   "FRK_ConfigAppend"(Scope := #Scope,
                      Item := 'CatalogCount',
                      ValueText := WSTRING#'0',
                      ValueType := 0,
                      ReadLevel := #ReadLevel,
                      Readable := #Readable,
                      Cursor := #Cursor,
                      Page := #Page);
   "FRK_ConfigAppend"(Scope := #Scope,
                      Item := 'AvailableModelCount',
                      ValueText := INT_TO_WSTRING(#ModelCount),
                      ValueType := 0,
                      ReadLevel := #ReadLevel,
                      Readable := #Readable,
                      Cursor := #Cursor,
                      Page := #Page);
   FOR #Index := 0 TO 6 DO
       #IndexText := INT_TO_STRING(#Index);
       IF #IndexText[1] = '+' THEN
           #IndexText := DELETE(IN := #IndexText, L := 1, P := 1);
       END_IF;
       #Prefix := CONCAT(IN1 := 'ModePolicy/ModePolicy[', IN2 := #IndexText);
       #Prefix := CONCAT(IN1 := #Prefix, IN2 := ']/');
       #Item := CONCAT(IN1 := #Prefix, IN2 := 'Shield');
       "FRK_ConfigAppend"(Scope := #Scope,
                          Item := #Item,
                          ValueText := STRING_TO_WSTRING(DINT_TO_STRING(#Policy[#Index].Shield)),
                          ValueType := 0,
                          ReadLevel := #ReadLevel,
                          Readable := #Readable,
                          Cursor := #Cursor,
                          Page := #Page);
       #Item := CONCAT(IN1 := #Prefix, IN2 := 'Style');
       "FRK_ConfigAppend"(Scope := #Scope,
                          Item := #Item,
                          ValueText := STRING_TO_WSTRING(DINT_TO_STRING(#Policy[#Index].Style)),
                          ValueType := 0,
                          ReadLevel := #ReadLevel,
                          Readable := #Readable,
                          Cursor := #Cursor,
                          Page := #Page);
   END_FOR;
END_FUNCTION

FUNCTION "FRK_Config_DeclarationCell" : Void   // FC141, SCL
{ S7_Optimized_Access := 'TRUE' }
VERSION : 0.1
// stored: AutoNumber true, IsIECCheckEnabled false, SetENOAutomatically false, UDAEnableTagReadback false
   VAR_INPUT
      Access : "FRK_Access";
      RootIndex : Int;
      ModelIndex : UDInt;
   END_VAR
   VAR_IN_OUT
      Module : "FB_DeclarationCell";
      Cursor : "FRK_ConfigCursor";
      Page : "ST_ConfigPage";
   END_VAR
   VAR_TEMP
      Ok : Bool;
   END_VAR
BEGIN

   IF #ModelIndex = 0 THEN
       "FRK_ConfigCatalog"(Scope := #Module.Status.Name,
                           Catalog := #Module.Catalog,
                           Count := #Module.CatalogCount,
                           ReadLevel := #Access.Policy.Required[0],
                           Readable := #Access.CurrentLevel >= #Access.Policy.Required[0],
                           Cursor := #Cursor,
                           Page := #Page);
   END_IF;
   IF #ModelIndex = 0 THEN
       "FRK_CfgDef_DeclarationCell"(FieldIndex := 1);
       "FRK_ConfigScratch".Entry.Scope := STRING_TO_WSTRING(#Module.Status.Name);
       "FRK_ConfigScratch".Entry.ReadLevel := MAX(IN1 := #Access.Policy.Required[0], IN2 := "FRK_ConfigScratch".MinRead);
       "FRK_ConfigScratch".Entry.WriteLevel := MAX(IN1 := #Access.Policy.Required[1], IN2 := "FRK_ConfigScratch".MinWrite);
       "FRK_ConfigScratch".Entry.Readable := #Access.CurrentLevel >= "FRK_ConfigScratch".Entry.ReadLevel;
       "FRK_ConfigScratch".Entry.ModelScoped := FALSE;
       "FRK_ConfigScratch".Entry.ValueText := DINT_TO_WSTRING(TIME_TO_DINT(#Module.ParCfg.Timeout));
       IF NOT "FRK_ConfigScratch".Entry.Readable THEN
           "FRK_ConfigScratch".Entry.ValueText := WSTRING#'';
       END_IF;
       "FRK_ConfigAppendEntry"(Cursor := #Cursor,
                               Page := #Page);
   END_IF;
   IF #ModelIndex = 0 THEN
       "FRK_CfgDef_DeclarationCell"(FieldIndex := 2);
       "FRK_ConfigScratch".Entry.Scope := STRING_TO_WSTRING(#Module.Status.Name);
       "FRK_ConfigScratch".Entry.ReadLevel := MAX(IN1 := #Access.Policy.Required[0], IN2 := "FRK_ConfigScratch".MinRead);
       "FRK_ConfigScratch".Entry.WriteLevel := MAX(IN1 := #Access.Policy.Required[1], IN2 := "FRK_ConfigScratch".MinWrite);
       "FRK_ConfigScratch".Entry.Readable := #Access.CurrentLevel >= "FRK_ConfigScratch".Entry.ReadLevel;
       "FRK_ConfigScratch".Entry.ModelScoped := FALSE;
       "FRK_ConfigScratch".Entry.ValueText := DINT_TO_WSTRING(#Module.ParCfg.Preset);
       IF NOT "FRK_ConfigScratch".Entry.Readable THEN
           "FRK_ConfigScratch".Entry.ValueText := WSTRING#'';
       END_IF;
       "FRK_ConfigAppendEntry"(Cursor := #Cursor,
                               Page := #Page);
   END_IF;
   IF #ModelIndex = 0 THEN
       "FRK_Config_DeclarationCylinder"(Module := #Module.Clamp,
                                        Access := #Access,
                                        RootIndex := #RootIndex,
                                        ModelIndex := #ModelIndex,
                                        Cursor := #Cursor,
                                        Page := #Page);
   END_IF;
   IF #ModelIndex = 0 THEN
       "FRK_Config_DeclarationCylinder"(Module := #Module.Gate,
                                        Access := #Access,
                                        RootIndex := #RootIndex,
                                        ModelIndex := #ModelIndex,
                                        Cursor := #Cursor,
                                        Page := #Page);
   END_IF;
END_FUNCTION

FUNCTION "FRK_Config_DeclarationCylinder" : Void   // FC133, SCL
{ S7_Optimized_Access := 'TRUE' }
VERSION : 0.1
// stored: AutoNumber true, IsIECCheckEnabled false, SetENOAutomatically false, UDAEnableTagReadback false
   VAR_INPUT
      Access : "FRK_Access";
      RootIndex : Int;
      ModelIndex : UDInt;
   END_VAR
   VAR_IN_OUT
      Module : "FB_DeclarationCylinder";
      Cursor : "FRK_ConfigCursor";
      Page : "ST_ConfigPage";
   END_VAR
   VAR_TEMP
      Ok : Bool;
   END_VAR
BEGIN

   IF #ModelIndex = 0 THEN
       "FRK_ConfigCatalog"(Scope := #Module.Status.Name,
                           Catalog := #Module.Catalog,
                           Count := #Module.CatalogCount,
                           ReadLevel := #Access.Policy.Required[0],
                           Readable := #Access.CurrentLevel >= #Access.Policy.Required[0],
                           Cursor := #Cursor,
                           Page := #Page);
   END_IF;
   IF #ModelIndex = 0 THEN
       "FRK_CfgDef_DeclarationCylinder"(FieldIndex := 1);
       "FRK_ConfigScratch".Entry.Scope := STRING_TO_WSTRING(#Module.Status.Name);
       "FRK_ConfigScratch".Entry.ReadLevel := MAX(IN1 := #Access.Policy.Required[0], IN2 := "FRK_ConfigScratch".MinRead);
       "FRK_ConfigScratch".Entry.WriteLevel := MAX(IN1 := #Access.Policy.Required[1], IN2 := "FRK_ConfigScratch".MinWrite);
       "FRK_ConfigScratch".Entry.Readable := #Access.CurrentLevel >= "FRK_ConfigScratch".Entry.ReadLevel;
       "FRK_ConfigScratch".Entry.ModelScoped := FALSE;
       "FRK_ConfigScratch".Entry.ValueText := DINT_TO_WSTRING(TIME_TO_DINT(#Module.ParCfg.Timeout));
       IF NOT "FRK_ConfigScratch".Entry.Readable THEN
           "FRK_ConfigScratch".Entry.ValueText := WSTRING#'';
       END_IF;
       "FRK_ConfigAppendEntry"(Cursor := #Cursor,
                               Page := #Page);
   END_IF;
   IF #ModelIndex = 0 THEN
       "FRK_CfgDef_DeclarationCylinder"(FieldIndex := 2);
       "FRK_ConfigScratch".Entry.Scope := STRING_TO_WSTRING(#Module.Status.Name);
       "FRK_ConfigScratch".Entry.ReadLevel := MAX(IN1 := #Access.Policy.Required[0], IN2 := "FRK_ConfigScratch".MinRead);
       "FRK_ConfigScratch".Entry.WriteLevel := MAX(IN1 := #Access.Policy.Required[1], IN2 := "FRK_ConfigScratch".MinWrite);
       "FRK_ConfigScratch".Entry.Readable := #Access.CurrentLevel >= "FRK_ConfigScratch".Entry.ReadLevel;
       "FRK_ConfigScratch".Entry.ModelScoped := FALSE;
       "FRK_ConfigScratch".Entry.ValueText := DINT_TO_WSTRING(#Module.ParCfg.Preset);
       IF NOT "FRK_ConfigScratch".Entry.Readable THEN
           "FRK_ConfigScratch".Entry.ValueText := WSTRING#'';
       END_IF;
       "FRK_ConfigAppendEntry"(Cursor := #Cursor,
                               Page := #Page);
   END_IF;
END_FUNCTION

FUNCTION "FRK_Config_DeclarationUnit" : Void   // FC166, SCL
{ S7_Optimized_Access := 'TRUE' }
VERSION : 0.1
// stored: AutoNumber true, IsIECCheckEnabled false, SetENOAutomatically false, UDAEnableTagReadback false
   VAR_INPUT
      Access : "FRK_Access";
      RootIndex : Int;
      ModelIndex : UDInt;
   END_VAR
   VAR_IN_OUT
      Core : "FRK_Core";
      Status : "ST_ModuleStatus";
      ParCfg : "ST_DeclarationParCfg";
      ModePolicy : Array[0..6] of "ST_ModePolicy";
      AvailableModelCount : Int;
      StationCfg : "ST_UnitProbeStationCfg";
      Cell : "FB_DeclarationCell";
      Satellite : "FB_SatelliteUnit";
      Cursor : "FRK_ConfigCursor";
      Page : "ST_ConfigPage";
   END_VAR
   VAR_TEMP
      Ok : Bool;
   END_VAR
BEGIN

   IF #ModelIndex = 0 THEN
       "FRK_ConfigUnit"(Scope := #Status.Name,
                        Policy := #ModePolicy,
                        ModelCount := #AvailableModelCount,
                        ReadLevel := #Access.Policy.Required[0],
                        Readable := #Access.CurrentLevel >= #Access.Policy.Required[0],
                        Cursor := #Cursor,
                        Page := #Page);
   END_IF;
   IF #ModelIndex = 0 THEN
       "FRK_ConfigAppend"(Scope := #Status.Name,
                          Item := 'AvailableModels/AvailableModels[1]/ModelCode',
                          ValueText := WSTRING#'MODEL_A',
                          ValueType := 1,
                          ReadLevel := #Access.Policy.Required[0],
                          Readable := #Access.CurrentLevel >= #Access.Policy.Required[0],
                          Cursor := #Cursor,
                          Page := #Page);
       "FRK_ConfigAppend"(Scope := #Status.Name,
                          Item := 'AvailableModels/AvailableModels[2]/ModelCode',
                          ValueText := WSTRING#'MODEL_B',
                          ValueType := 1,
                          ReadLevel := #Access.Policy.Required[0],
                          Readable := #Access.CurrentLevel >= #Access.Policy.Required[0],
                          Cursor := #Cursor,
                          Page := #Page);
   END_IF;
   IF (#ModelIndex = 0 OR #Core.ParentIndex = 0) THEN
       "FRK_CfgDef_DeclarationUnit"(FieldIndex := 1);
       "FRK_ConfigScratch".Entry.Scope := STRING_TO_WSTRING(#Status.Name);
       "FRK_ConfigScratch".Entry.ReadLevel := MAX(IN1 := #Access.Policy.Required[0], IN2 := "FRK_ConfigScratch".MinRead);
       "FRK_ConfigScratch".Entry.WriteLevel := MAX(IN1 := #Access.Policy.Required[1], IN2 := "FRK_ConfigScratch".MinWrite);
       "FRK_ConfigScratch".Entry.Readable := #Access.CurrentLevel >= "FRK_ConfigScratch".Entry.ReadLevel;
       "FRK_ConfigScratch".Entry.ModelScoped := #Core.ParentIndex = 0;
       IF #ModelIndex <> 0 THEN
           "FRK_ConfigScratch".Entry.RequiresReady := "FRK_ConfigScratch".Entry.RequiresReady AND "FRK_ConfigModelCode"(RootIndex := #RootIndex, ModelIndex := #ModelIndex) = "FRK_ConfigStore".ActiveModels[#RootIndex];
           #Ok := "FRK_ConfigGet"(Scope := #Status.Name, ModelCode := "FRK_ConfigModelCode"(RootIndex := #RootIndex, ModelIndex := #ModelIndex));
           IF NOT #Ok THEN
               "FRK_ConfigScratch".Entry.Readable := FALSE;
           END_IF;
       ELSE
           "FRK_ConfigScratch".Entry.ValueText := DINT_TO_WSTRING(TIME_TO_DINT(#ParCfg.Timeout));
       END_IF;
       IF NOT "FRK_ConfigScratch".Entry.Readable THEN
           "FRK_ConfigScratch".Entry.ValueText := WSTRING#'';
       END_IF;
       "FRK_ConfigAppendEntry"(Cursor := #Cursor,
                               Page := #Page);
   END_IF;
   IF (#ModelIndex = 0 OR #Core.ParentIndex = 0) THEN
       "FRK_CfgDef_DeclarationUnit"(FieldIndex := 2);
       "FRK_ConfigScratch".Entry.Scope := STRING_TO_WSTRING(#Status.Name);
       "FRK_ConfigScratch".Entry.ReadLevel := MAX(IN1 := #Access.Policy.Required[0], IN2 := "FRK_ConfigScratch".MinRead);
       "FRK_ConfigScratch".Entry.WriteLevel := MAX(IN1 := #Access.Policy.Required[1], IN2 := "FRK_ConfigScratch".MinWrite);
       "FRK_ConfigScratch".Entry.Readable := #Access.CurrentLevel >= "FRK_ConfigScratch".Entry.ReadLevel;
       "FRK_ConfigScratch".Entry.ModelScoped := #Core.ParentIndex = 0;
       IF #ModelIndex <> 0 THEN
           "FRK_ConfigScratch".Entry.RequiresReady := "FRK_ConfigScratch".Entry.RequiresReady AND "FRK_ConfigModelCode"(RootIndex := #RootIndex, ModelIndex := #ModelIndex) = "FRK_ConfigStore".ActiveModels[#RootIndex];
           #Ok := "FRK_ConfigGet"(Scope := #Status.Name, ModelCode := "FRK_ConfigModelCode"(RootIndex := #RootIndex, ModelIndex := #ModelIndex));
           IF NOT #Ok THEN
               "FRK_ConfigScratch".Entry.Readable := FALSE;
           END_IF;
       ELSE
           "FRK_ConfigScratch".Entry.ValueText := DINT_TO_WSTRING(#ParCfg.Preset);
       END_IF;
       IF NOT "FRK_ConfigScratch".Entry.Readable THEN
           "FRK_ConfigScratch".Entry.ValueText := WSTRING#'';
       END_IF;
       "FRK_ConfigAppendEntry"(Cursor := #Cursor,
                               Page := #Page);
   END_IF;
   IF #ModelIndex = 0 THEN
       "FRK_CfgDef_DeclarationUnit"(FieldIndex := 3);
       "FRK_ConfigScratch".Entry.Scope := STRING_TO_WSTRING(#Status.Name);
       "FRK_ConfigScratch".Entry.ReadLevel := MAX(IN1 := #Access.Policy.Required[0], IN2 := "FRK_ConfigScratch".MinRead);
       "FRK_ConfigScratch".Entry.WriteLevel := MAX(IN1 := #Access.Policy.Required[1], IN2 := "FRK_ConfigScratch".MinWrite);
       "FRK_ConfigScratch".Entry.Readable := #Access.CurrentLevel >= "FRK_ConfigScratch".Entry.ReadLevel;
       "FRK_ConfigScratch".Entry.ModelScoped := FALSE;
       "FRK_ConfigScratch".Entry.ValueText := STRING_TO_WSTRING(#StationCfg.SiteLabel);
       IF NOT "FRK_ConfigScratch".Entry.Readable THEN
           "FRK_ConfigScratch".Entry.ValueText := WSTRING#'';
       END_IF;
       "FRK_ConfigAppendEntry"(Cursor := #Cursor,
                               Page := #Page);
   END_IF;
   IF #ModelIndex = 0 THEN
       "FRK_CfgDef_DeclarationUnit"(FieldIndex := 4);
       "FRK_ConfigScratch".Entry.Scope := STRING_TO_WSTRING(#Status.Name);
       "FRK_ConfigScratch".Entry.ReadLevel := MAX(IN1 := #Access.Policy.Required[0], IN2 := "FRK_ConfigScratch".MinRead);
       "FRK_ConfigScratch".Entry.WriteLevel := MAX(IN1 := #Access.Policy.Required[1], IN2 := "FRK_ConfigScratch".MinWrite);
       "FRK_ConfigScratch".Entry.Readable := #Access.CurrentLevel >= "FRK_ConfigScratch".Entry.ReadLevel;
       "FRK_ConfigScratch".Entry.ModelScoped := FALSE;
       "FRK_ConfigScratch".Entry.ValueText := STRING_TO_WSTRING(#StationCfg.LongText);
       IF NOT "FRK_ConfigScratch".Entry.Readable THEN
           "FRK_ConfigScratch".Entry.ValueText := WSTRING#'';
       END_IF;
       "FRK_ConfigAppendEntry"(Cursor := #Cursor,
                               Page := #Page);
   END_IF;
   IF #ModelIndex = 0 THEN
       "FRK_CfgDef_DeclarationUnit"(FieldIndex := 5);
       "FRK_ConfigScratch".Entry.Scope := STRING_TO_WSTRING(#Status.Name);
       "FRK_ConfigScratch".Entry.ReadLevel := MAX(IN1 := #Access.Policy.Required[0], IN2 := "FRK_ConfigScratch".MinRead);
       "FRK_ConfigScratch".Entry.WriteLevel := MAX(IN1 := #Access.Policy.Required[1], IN2 := "FRK_ConfigScratch".MinWrite);
       "FRK_ConfigScratch".Entry.Readable := #Access.CurrentLevel >= "FRK_ConfigScratch".Entry.ReadLevel;
       "FRK_ConfigScratch".Entry.ModelScoped := FALSE;
       IF #StationCfg.Enabled THEN
           "FRK_ConfigScratch".Entry.ValueText := WSTRING#'true';
       ELSE
           "FRK_ConfigScratch".Entry.ValueText := WSTRING#'false';
       END_IF;
       IF NOT "FRK_ConfigScratch".Entry.Readable THEN
           "FRK_ConfigScratch".Entry.ValueText := WSTRING#'';
       END_IF;
       "FRK_ConfigAppendEntry"(Cursor := #Cursor,
                               Page := #Page);
   END_IF;
   IF #ModelIndex = 0 THEN
       "FRK_Config_DeclarationCell"(Module := #Cell,
                                    Access := #Access,
                                    RootIndex := #RootIndex,
                                    ModelIndex := #ModelIndex,
                                    Cursor := #Cursor,
                                    Page := #Page);
   END_IF;
   IF #ModelIndex = 0 THEN
       "FRK_Config_SatelliteUnit"(Module := #Satellite,
                                  Access := #Access,
                                  RootIndex := #RootIndex,
                                  ModelIndex := #ModelIndex,
                                  Cursor := #Cursor,
                                  Page := #Page);
   END_IF;
END_FUNCTION

FUNCTION "FRK_Config_InnerUnit" : Void   // FC150, SCL
{ S7_Optimized_Access := 'TRUE' }
VERSION : 0.1
// stored: AutoNumber true, IsIECCheckEnabled false, SetENOAutomatically false, UDAEnableTagReadback false
   VAR_INPUT
      Access : "FRK_Access";
      RootIndex : Int;
      ModelIndex : UDInt;
   END_VAR
   VAR_IN_OUT
      Module : "FB_InnerUnit";
      Cursor : "FRK_ConfigCursor";
      Page : "ST_ConfigPage";
   END_VAR
   VAR_TEMP
      Ok : Bool;
   END_VAR
BEGIN

   IF #ModelIndex = 0 THEN
       "FRK_ConfigUnit"(Scope := #Module.Status.Name,
                        Policy := #Module.ModePolicy,
                        ModelCount := 0,
                        ReadLevel := #Access.Policy.Required[0],
                        Readable := #Access.CurrentLevel >= #Access.Policy.Required[0],
                        Cursor := #Cursor,
                        Page := #Page);
   END_IF;
   IF #ModelIndex = 0 THEN
       "FRK_CfgDef_InnerUnit"(FieldIndex := 1);
       "FRK_ConfigScratch".Entry.Scope := STRING_TO_WSTRING(#Module.Status.Name);
       "FRK_ConfigScratch".Entry.ReadLevel := MAX(IN1 := #Access.Policy.Required[0], IN2 := "FRK_ConfigScratch".MinRead);
       "FRK_ConfigScratch".Entry.WriteLevel := MAX(IN1 := #Access.Policy.Required[1], IN2 := "FRK_ConfigScratch".MinWrite);
       "FRK_ConfigScratch".Entry.Readable := #Access.CurrentLevel >= "FRK_ConfigScratch".Entry.ReadLevel;
       "FRK_ConfigScratch".Entry.ModelScoped := FALSE;
       "FRK_ConfigScratch".Entry.ValueText := DINT_TO_WSTRING(TIME_TO_DINT(#Module.ParCfg.Timeout));
       IF NOT "FRK_ConfigScratch".Entry.Readable THEN
           "FRK_ConfigScratch".Entry.ValueText := WSTRING#'';
       END_IF;
       "FRK_ConfigAppendEntry"(Cursor := #Cursor,
                               Page := #Page);
   END_IF;
   IF #ModelIndex = 0 THEN
       "FRK_CfgDef_InnerUnit"(FieldIndex := 2);
       "FRK_ConfigScratch".Entry.Scope := STRING_TO_WSTRING(#Module.Status.Name);
       "FRK_ConfigScratch".Entry.ReadLevel := MAX(IN1 := #Access.Policy.Required[0], IN2 := "FRK_ConfigScratch".MinRead);
       "FRK_ConfigScratch".Entry.WriteLevel := MAX(IN1 := #Access.Policy.Required[1], IN2 := "FRK_ConfigScratch".MinWrite);
       "FRK_ConfigScratch".Entry.Readable := #Access.CurrentLevel >= "FRK_ConfigScratch".Entry.ReadLevel;
       "FRK_ConfigScratch".Entry.ModelScoped := FALSE;
       "FRK_ConfigScratch".Entry.ValueText := DINT_TO_WSTRING(#Module.ParCfg.Preset);
       IF NOT "FRK_ConfigScratch".Entry.Readable THEN
           "FRK_ConfigScratch".Entry.ValueText := WSTRING#'';
       END_IF;
       "FRK_ConfigAppendEntry"(Cursor := #Cursor,
                               Page := #Page);
   END_IF;
   IF #ModelIndex = 0 THEN
       "FRK_CfgDef_InnerUnit"(FieldIndex := 3);
       "FRK_ConfigScratch".Entry.Scope := STRING_TO_WSTRING(#Module.Status.Name);
       "FRK_ConfigScratch".Entry.ReadLevel := MAX(IN1 := #Access.Policy.Required[0], IN2 := "FRK_ConfigScratch".MinRead);
       "FRK_ConfigScratch".Entry.WriteLevel := MAX(IN1 := #Access.Policy.Required[1], IN2 := "FRK_ConfigScratch".MinWrite);
       "FRK_ConfigScratch".Entry.Readable := #Access.CurrentLevel >= "FRK_ConfigScratch".Entry.ReadLevel;
       "FRK_ConfigScratch".Entry.ModelScoped := FALSE;
       "FRK_ConfigScratch".Entry.ValueText := STRING_TO_WSTRING(#Module.StationCfg.SiteLabel);
       IF NOT "FRK_ConfigScratch".Entry.Readable THEN
           "FRK_ConfigScratch".Entry.ValueText := WSTRING#'';
       END_IF;
       "FRK_ConfigAppendEntry"(Cursor := #Cursor,
                               Page := #Page);
   END_IF;
   IF #ModelIndex = 0 THEN
       "FRK_CfgDef_InnerUnit"(FieldIndex := 4);
       "FRK_ConfigScratch".Entry.Scope := STRING_TO_WSTRING(#Module.Status.Name);
       "FRK_ConfigScratch".Entry.ReadLevel := MAX(IN1 := #Access.Policy.Required[0], IN2 := "FRK_ConfigScratch".MinRead);
       "FRK_ConfigScratch".Entry.WriteLevel := MAX(IN1 := #Access.Policy.Required[1], IN2 := "FRK_ConfigScratch".MinWrite);
       "FRK_ConfigScratch".Entry.Readable := #Access.CurrentLevel >= "FRK_ConfigScratch".Entry.ReadLevel;
       "FRK_ConfigScratch".Entry.ModelScoped := FALSE;
       "FRK_ConfigScratch".Entry.ValueText := STRING_TO_WSTRING(#Module.StationCfg.LongText);
       IF NOT "FRK_ConfigScratch".Entry.Readable THEN
           "FRK_ConfigScratch".Entry.ValueText := WSTRING#'';
       END_IF;
       "FRK_ConfigAppendEntry"(Cursor := #Cursor,
                               Page := #Page);
   END_IF;
   IF #ModelIndex = 0 THEN
       "FRK_CfgDef_InnerUnit"(FieldIndex := 5);
       "FRK_ConfigScratch".Entry.Scope := STRING_TO_WSTRING(#Module.Status.Name);
       "FRK_ConfigScratch".Entry.ReadLevel := MAX(IN1 := #Access.Policy.Required[0], IN2 := "FRK_ConfigScratch".MinRead);
       "FRK_ConfigScratch".Entry.WriteLevel := MAX(IN1 := #Access.Policy.Required[1], IN2 := "FRK_ConfigScratch".MinWrite);
       "FRK_ConfigScratch".Entry.Readable := #Access.CurrentLevel >= "FRK_ConfigScratch".Entry.ReadLevel;
       "FRK_ConfigScratch".Entry.ModelScoped := FALSE;
       IF #Module.StationCfg.Enabled THEN
           "FRK_ConfigScratch".Entry.ValueText := WSTRING#'true';
       ELSE
           "FRK_ConfigScratch".Entry.ValueText := WSTRING#'false';
       END_IF;
       IF NOT "FRK_ConfigScratch".Entry.Readable THEN
           "FRK_ConfigScratch".Entry.ValueText := WSTRING#'';
       END_IF;
       "FRK_ConfigAppendEntry"(Cursor := #Cursor,
                               Page := #Page);
   END_IF;
   IF #ModelIndex = 0 THEN
       "FRK_Config_DeclarationCell"(Module := #Module.Cell,
                                    Access := #Access,
                                    RootIndex := #RootIndex,
                                    ModelIndex := #ModelIndex,
                                    Cursor := #Cursor,
                                    Page := #Page);
   END_IF;
END_FUNCTION

FUNCTION "FRK_Config_SatelliteUnit" : Void   // FC158, SCL
{ S7_Optimized_Access := 'TRUE' }
VERSION : 0.1
// stored: AutoNumber true, IsIECCheckEnabled false, SetENOAutomatically false, UDAEnableTagReadback false
   VAR_INPUT
      Access : "FRK_Access";
      RootIndex : Int;
      ModelIndex : UDInt;
   END_VAR
   VAR_IN_OUT
      Module : "FB_SatelliteUnit";
      Cursor : "FRK_ConfigCursor";
      Page : "ST_ConfigPage";
   END_VAR
   VAR_TEMP
      Ok : Bool;
   END_VAR
BEGIN

   IF #ModelIndex = 0 THEN
       "FRK_ConfigUnit"(Scope := #Module.Status.Name,
                        Policy := #Module.ModePolicy,
                        ModelCount := 0,
                        ReadLevel := #Access.Policy.Required[0],
                        Readable := #Access.CurrentLevel >= #Access.Policy.Required[0],
                        Cursor := #Cursor,
                        Page := #Page);
   END_IF;
   IF #ModelIndex = 0 THEN
       "FRK_CfgDef_SatelliteUnit"(FieldIndex := 1);
       "FRK_ConfigScratch".Entry.Scope := STRING_TO_WSTRING(#Module.Status.Name);
       "FRK_ConfigScratch".Entry.ReadLevel := MAX(IN1 := #Access.Policy.Required[0], IN2 := "FRK_ConfigScratch".MinRead);
       "FRK_ConfigScratch".Entry.WriteLevel := MAX(IN1 := #Access.Policy.Required[1], IN2 := "FRK_ConfigScratch".MinWrite);
       "FRK_ConfigScratch".Entry.Readable := #Access.CurrentLevel >= "FRK_ConfigScratch".Entry.ReadLevel;
       "FRK_ConfigScratch".Entry.ModelScoped := FALSE;
       "FRK_ConfigScratch".Entry.ValueText := DINT_TO_WSTRING(TIME_TO_DINT(#Module.ParCfg.Timeout));
       IF NOT "FRK_ConfigScratch".Entry.Readable THEN
           "FRK_ConfigScratch".Entry.ValueText := WSTRING#'';
       END_IF;
       "FRK_ConfigAppendEntry"(Cursor := #Cursor,
                               Page := #Page);
   END_IF;
   IF #ModelIndex = 0 THEN
       "FRK_CfgDef_SatelliteUnit"(FieldIndex := 2);
       "FRK_ConfigScratch".Entry.Scope := STRING_TO_WSTRING(#Module.Status.Name);
       "FRK_ConfigScratch".Entry.ReadLevel := MAX(IN1 := #Access.Policy.Required[0], IN2 := "FRK_ConfigScratch".MinRead);
       "FRK_ConfigScratch".Entry.WriteLevel := MAX(IN1 := #Access.Policy.Required[1], IN2 := "FRK_ConfigScratch".MinWrite);
       "FRK_ConfigScratch".Entry.Readable := #Access.CurrentLevel >= "FRK_ConfigScratch".Entry.ReadLevel;
       "FRK_ConfigScratch".Entry.ModelScoped := FALSE;
       "FRK_ConfigScratch".Entry.ValueText := DINT_TO_WSTRING(#Module.ParCfg.Preset);
       IF NOT "FRK_ConfigScratch".Entry.Readable THEN
           "FRK_ConfigScratch".Entry.ValueText := WSTRING#'';
       END_IF;
       "FRK_ConfigAppendEntry"(Cursor := #Cursor,
                               Page := #Page);
   END_IF;
   IF #ModelIndex = 0 THEN
       "FRK_CfgDef_SatelliteUnit"(FieldIndex := 3);
       "FRK_ConfigScratch".Entry.Scope := STRING_TO_WSTRING(#Module.Status.Name);
       "FRK_ConfigScratch".Entry.ReadLevel := MAX(IN1 := #Access.Policy.Required[0], IN2 := "FRK_ConfigScratch".MinRead);
       "FRK_ConfigScratch".Entry.WriteLevel := MAX(IN1 := #Access.Policy.Required[1], IN2 := "FRK_ConfigScratch".MinWrite);
       "FRK_ConfigScratch".Entry.Readable := #Access.CurrentLevel >= "FRK_ConfigScratch".Entry.ReadLevel;
       "FRK_ConfigScratch".Entry.ModelScoped := FALSE;
       "FRK_ConfigScratch".Entry.ValueText := STRING_TO_WSTRING(#Module.StationCfg.SiteLabel);
       IF NOT "FRK_ConfigScratch".Entry.Readable THEN
           "FRK_ConfigScratch".Entry.ValueText := WSTRING#'';
       END_IF;
       "FRK_ConfigAppendEntry"(Cursor := #Cursor,
                               Page := #Page);
   END_IF;
   IF #ModelIndex = 0 THEN
       "FRK_CfgDef_SatelliteUnit"(FieldIndex := 4);
       "FRK_ConfigScratch".Entry.Scope := STRING_TO_WSTRING(#Module.Status.Name);
       "FRK_ConfigScratch".Entry.ReadLevel := MAX(IN1 := #Access.Policy.Required[0], IN2 := "FRK_ConfigScratch".MinRead);
       "FRK_ConfigScratch".Entry.WriteLevel := MAX(IN1 := #Access.Policy.Required[1], IN2 := "FRK_ConfigScratch".MinWrite);
       "FRK_ConfigScratch".Entry.Readable := #Access.CurrentLevel >= "FRK_ConfigScratch".Entry.ReadLevel;
       "FRK_ConfigScratch".Entry.ModelScoped := FALSE;
       "FRK_ConfigScratch".Entry.ValueText := STRING_TO_WSTRING(#Module.StationCfg.LongText);
       IF NOT "FRK_ConfigScratch".Entry.Readable THEN
           "FRK_ConfigScratch".Entry.ValueText := WSTRING#'';
       END_IF;
       "FRK_ConfigAppendEntry"(Cursor := #Cursor,
                               Page := #Page);
   END_IF;
   IF #ModelIndex = 0 THEN
       "FRK_CfgDef_SatelliteUnit"(FieldIndex := 5);
       "FRK_ConfigScratch".Entry.Scope := STRING_TO_WSTRING(#Module.Status.Name);
       "FRK_ConfigScratch".Entry.ReadLevel := MAX(IN1 := #Access.Policy.Required[0], IN2 := "FRK_ConfigScratch".MinRead);
       "FRK_ConfigScratch".Entry.WriteLevel := MAX(IN1 := #Access.Policy.Required[1], IN2 := "FRK_ConfigScratch".MinWrite);
       "FRK_ConfigScratch".Entry.Readable := #Access.CurrentLevel >= "FRK_ConfigScratch".Entry.ReadLevel;
       "FRK_ConfigScratch".Entry.ModelScoped := FALSE;
       IF #Module.StationCfg.Enabled THEN
           "FRK_ConfigScratch".Entry.ValueText := WSTRING#'true';
       ELSE
           "FRK_ConfigScratch".Entry.ValueText := WSTRING#'false';
       END_IF;
       IF NOT "FRK_ConfigScratch".Entry.Readable THEN
           "FRK_ConfigScratch".Entry.ValueText := WSTRING#'';
       END_IF;
       "FRK_ConfigAppendEntry"(Cursor := #Cursor,
                               Page := #Page);
   END_IF;
   IF #ModelIndex = 0 THEN
       "FRK_Config_DeclarationCell"(Module := #Module.Cell,
                                    Access := #Access,
                                    RootIndex := #RootIndex,
                                    ModelIndex := #ModelIndex,
                                    Cursor := #Cursor,
                                    Page := #Page);
   END_IF;
   IF #ModelIndex = 0 THEN
       "FRK_Config_InnerUnit"(Module := #Module.Inner,
                              Access := #Access,
                              RootIndex := #RootIndex,
                              ModelIndex := #ModelIndex,
                              Cursor := #Cursor,
                              Page := #Page);
   END_IF;
END_FUNCTION

FUNCTION "FRK_CrcByte" : DWord   // FC56, SCL
{ S7_Optimized_Access := 'TRUE' }
VERSION : 0.1
// Reference-1500 LOCAL_RETAIN adapter. No sessions or plaintext credentials.
//  CRC-32 arithmetic comes from Core F_Crc32; encoding is binding-local, versioned.
// stored: AutoNumber true, IsIECCheckEnabled false, SetENOAutomatically false, UDAEnableTagReadback false
   VAR_INPUT
      Previous : DWord;
      Value : Byte;
   END_VAR
   VAR_TEMP
      BitIndex : Int;
      Work : DWord;
   END_VAR
BEGIN

   #Work := #Previous XOR BYTE_TO_DWORD(#Value);
   FOR #BitIndex := 0 TO 7 DO
       IF (#Work AND DWORD#1) <> 0 THEN
           #Work := SHR(IN := #Work, N := 1) XOR DWORD#16#EDB88320;
       ELSE
           #Work := SHR(IN := #Work, N := 1);
       END_IF;
   END_FOR;
   #FRK_CrcByte := #Work;
END_FUNCTION

FUNCTION "FRK_CrcNumber" : DWord   // FC57, SCL
{ S7_Optimized_Access := 'TRUE' }
VERSION : 0.1
// stored: AutoNumber true, IsIECCheckEnabled false, SetENOAutomatically false, UDAEnableTagReadback false
   VAR_INPUT
      Previous : DWord;
      Value : UDInt;
   END_VAR
   VAR_TEMP
      Index : Int;
      Work : DWord;
   END_VAR
BEGIN

   #Work := #Previous;
   FOR #Index := 0 TO 3 DO
       #Work := "FRK_CrcByte"(Previous := #Work, Value := DWORD_TO_BYTE(SHR(IN := UDINT_TO_DWORD(#Value), N := INT_TO_UINT(#Index * 8))));
   END_FOR;
   #FRK_CrcNumber := #Work;
END_FUNCTION

FUNCTION "FRK_DecisionAsk" : Bool   // FC97, SCL
{ S7_Optimized_Access := 'TRUE' }
VERSION : 0.1
// stored: AutoNumber true, IsIECCheckEnabled false, SetENOAutomatically false, UDAEnableTagReadback false
   VAR_INPUT
      Owner : DInt;
      OwnerPath : WString;
      Request : "ST_DecisionRequest";
   END_VAR
   VAR_IN_OUT
      AlarmLog : "FRK_AlarmLog";
   END_VAR
   VAR_TEMP
      Candidate : "ST_DecisionRequest";
      Slot : Int;
      Index : Int;
      SameRequest : Bool;
      HasOption : Bool;
   END_VAR
BEGIN

   #FRK_DecisionAsk := FALSE;
   #Slot := "FRK_DecisionRoot"(Owner := #Owner, Create := TRUE);
   IF #Slot = 0 THEN
       RETURN;
   END_IF;
   #Candidate := #Request;
   IF #Candidate.SourcePath = WSTRING#'' THEN
       #Candidate.SourcePath := #OwnerPath;
   END_IF;
   IF "FRK_Decisions".Slots[#Slot].Request.Prompt <> WSTRING#'' THEN
       #SameRequest := "FRK_Decisions".Slots[#Slot].Owner = #Owner
       AND "FRK_Decisions".Slots[#Slot].Request.Prompt = #Candidate.Prompt
       AND "FRK_Decisions".Slots[#Slot].Request.SourcePath = #Candidate.SourcePath
       AND "FRK_Decisions".Slots[#Slot].Request.Default = #Candidate.Default
       AND "FRK_Decisions".Slots[#Slot].Request.Timeout = #Candidate.Timeout;
       FOR #Index := 1 TO 6 DO
           #SameRequest := #SameRequest AND "FRK_Decisions".Slots[#Slot].Request.Options[#Index] = #Candidate.Options[#Index];
       END_FOR;
       IF #SameRequest THEN
           #FRK_DecisionAsk := TRUE;
           RETURN;
       END_IF;
       IF NOT "FRK_Decisions".Slots[#Slot].OverlapLogged THEN
           "FRK_DecisionAudit"(AlarmLog := #AlarmLog,
                               Key := WSTRING#'std.audit.decisionOverlapRejected',
                               SourcePath := #Candidate.SourcePath,
                               Option := 0);
           "FRK_Decisions".Slots[#Slot].OverlapLogged := TRUE;
       END_IF;
       RETURN;
   END_IF;
   #HasOption := FALSE;
   FOR #Index := 1 TO 6 DO
       #HasOption := #HasOption OR #Candidate.Options[#Index] <> '';
   END_FOR;
   IF #Candidate.Prompt = WSTRING#'' OR #Candidate.Timeout < T#0ms OR NOT #HasOption
       OR #Candidate.SourcePath <> #OwnerPath OR #OwnerPath = WSTRING#'' THEN
       "FRK_DecisionAudit"(AlarmLog := #AlarmLog,
                           Key := WSTRING#'std.audit.decisionInvalidRejected',
                           SourcePath := #Candidate.SourcePath,
                           Option := #Candidate.Default);
       RETURN;
   END_IF;
   IF #Candidate.Timeout > T#0ms OR #Candidate.Default <> 0 THEN
       IF #Candidate.Default < 1 OR #Candidate.Default > 6 THEN
           "FRK_DecisionAudit"(AlarmLog := #AlarmLog,
                               Key := WSTRING#'std.audit.decisionInvalidRejected',
                               SourcePath := #Candidate.SourcePath,
                               Option := #Candidate.Default);
           RETURN;
       END_IF;
       IF #Candidate.Options[#Candidate.Default] = '' THEN
           "FRK_DecisionAudit"(AlarmLog := #AlarmLog,
                               Key := WSTRING#'std.audit.decisionInvalidRejected',
                               SourcePath := #Candidate.SourcePath,
                               Option := #Candidate.Default);
           RETURN;
       END_IF;
   END_IF;
   "FRK_Decisions".Slots[#Slot].Request := #Candidate;
   "FRK_Decisions".Slots[#Slot].Owner := #Owner;
   "FRK_Decisions".Slots[#Slot].AskedAt := "FRK_Clock".NowMs;
   "FRK_Decisions".Slots[#Slot].Answer := 0;
   "FRK_Decisions".Slots[#Slot].ResolutionLogged := FALSE;
   "FRK_Decisions".Slots[#Slot].OverlapLogged := FALSE;
   "FRK_DecisionAudit"(AlarmLog := #AlarmLog,
                       Key := WSTRING#'std.audit.decisionRequested',
                       SourcePath := #Candidate.SourcePath,
                       Option := 0);
   #FRK_DecisionAsk := TRUE;
END_FUNCTION

FUNCTION "FRK_DecisionAudit" : Void   // FC95, SCL
{ S7_Optimized_Access := 'TRUE' }
VERSION : 0.1
// stored: AutoNumber true, IsIECCheckEnabled false, SetENOAutomatically false, UDAEnableTagReadback false
   VAR_INPUT
      Key : WString;
      SourcePath : WString;
      Option : Int;
   END_VAR
   VAR_IN_OUT
      AlarmLog : "FRK_AlarmLog";
   END_VAR
   VAR_TEMP
      Diag : "ST_Diagnostic";
      Slot : Int;
      Gone : Bool;
   END_VAR
BEGIN

   #Diag := "FRK_UnitScratch".EmptyDiagnostic;
   #Diag.Description := #Key;
   IF #Option <> 0 THEN
       #Diag.Description := CONCAT(IN1 := #Diag.Description, IN2 := WSTRING#' option=');
       #Diag.Description := CONCAT(IN1 := #Diag.Description, IN2 := STRING_TO_WSTRING(INT_TO_STRING(#Option)));
   END_IF;
   #Diag.SourcePath := #SourcePath;
   #Diag.Severity := 0;
   #Diag.Category := 0;
   #Slot := "FRK_AlarmRaise"(AlarmLog := #AlarmLog, Diag := #Diag, ResetClass := 0);
   IF #Slot > 0 THEN
       #Gone := "FRK_AlarmGone"(AlarmLog := #AlarmLog, Slot := #Slot);
   END_IF;
END_FUNCTION

FUNCTION "FRK_DecisionClear" : Void   // FC96, SCL
{ S7_Optimized_Access := 'TRUE' }
VERSION : 0.1
// stored: AutoNumber true, IsIECCheckEnabled false, SetENOAutomatically false, UDAEnableTagReadback false
   VAR_IN_OUT
      Slot : "FRK_DecisionSlot";
   END_VAR
   VAR_TEMP
      Index : Int;
   END_VAR
BEGIN

   #Slot.Request.Prompt := WSTRING#'';
   #Slot.Request.SourcePath := WSTRING#'';
   #Slot.Request.Default := 0;
   #Slot.Request.Timeout := T#0ms;
   FOR #Index := 1 TO 6 DO
       #Slot.Request.Options[#Index] := '';
   END_FOR;
   #Slot.Answer := 0;
   #Slot.Owner := 0;
   #Slot.OverlapLogged := FALSE;
   #Slot.ResolutionLogged := FALSE;
END_FUNCTION

FUNCTION "FRK_DecisionCyclic" : Void   // FC99, SCL
{ S7_Optimized_Access := 'TRUE' }
VERSION : 0.1
// stored: AutoNumber true, IsIECCheckEnabled false, SetENOAutomatically false, UDAEnableTagReadback false
   VAR_INPUT
      Owner : DInt;
      Busy : Bool;
      Reset : Bool;
   END_VAR
   VAR_IN_OUT
      AlarmLog : "FRK_AlarmLog";
   END_VAR
   VAR_TEMP
      Slot : Int;
      Elapsed : UDInt;
   END_VAR
BEGIN

   IF #Owner < 1 OR #Owner > "FRK_Registry".Count THEN
       RETURN;
   END_IF;
   // Only the root resolves/withdraws its slot; an idle nested Unit cannot
   // cancel a root's running decision.
   IF "FRK_Registry".Rows[#Owner].Parent <> 0 THEN
       RETURN;
   END_IF;
   #Slot := "FRK_DecisionRoot"(Owner := #Owner, Create := FALSE);
   IF #Slot = 0 THEN
       RETURN;
   END_IF;
   IF "FRK_Decisions".Slots[#Slot].Request.Prompt = WSTRING#'' THEN
       RETURN;
   END_IF;
   IF #Reset OR NOT #Busy THEN
       "FRK_DecisionAudit"(AlarmLog := #AlarmLog,
                           Key := WSTRING#'std.audit.decisionWithdrawn',
                           SourcePath := "FRK_Decisions".Slots[#Slot].Request.SourcePath,
                           Option := 0);
       "FRK_DecisionClear"(Slot := "FRK_Decisions".Slots[#Slot]);
       RETURN;
   END_IF;
   IF "FRK_Decisions".Slots[#Slot].Answer <> 0 THEN
       IF NOT "FRK_Decisions".Slots[#Slot].ResolutionLogged THEN
           "FRK_DecisionAudit"(AlarmLog := #AlarmLog,
                               Key := WSTRING#'std.audit.decisionOperatorResolved',
                               SourcePath := "FRK_Decisions".Slots[#Slot].Request.SourcePath,
                               Option := "FRK_Decisions".Slots[#Slot].Answer);
           "FRK_Decisions".Slots[#Slot].ResolutionLogged := TRUE;
       END_IF;
       RETURN;
   END_IF;
   IF "FRK_Decisions".Slots[#Slot].Request.Timeout <= T#0ms THEN
       RETURN;
   END_IF;
   #Elapsed := "FRK_Clock".NowMs - "FRK_Decisions".Slots[#Slot].AskedAt;
   IF #Elapsed >= DINT_TO_UDINT(TIME_TO_DINT("FRK_Decisions".Slots[#Slot].Request.Timeout)) THEN
       "FRK_Decisions".Slots[#Slot].Answer := "FRK_Decisions".Slots[#Slot].Request.Default;
       "FRK_DecisionAudit"(AlarmLog := #AlarmLog,
                           Key := WSTRING#'std.audit.decisionTimeoutResolved',
                           SourcePath := "FRK_Decisions".Slots[#Slot].Request.SourcePath,
                           Option := "FRK_Decisions".Slots[#Slot].Answer);
       "FRK_Decisions".Slots[#Slot].ResolutionLogged := TRUE;
   END_IF;
END_FUNCTION

FUNCTION "FRK_DecisionPublish" : Void   // FC101, SCL
{ S7_Optimized_Access := 'TRUE' }
VERSION : 0.1
// stored: AutoNumber true, IsIECCheckEnabled false, SetENOAutomatically false, UDAEnableTagReadback false
   VAR_INPUT
      Owner : DInt;
   END_VAR
   VAR_IN_OUT
      Decision : "ST_DecisionRequest";
      DecisionAnswer : Int;
   END_VAR
   VAR_TEMP
      Slot : Int;
   END_VAR
BEGIN

   #Slot := "FRK_DecisionRoot"(Owner := #Owner, Create := FALSE);
   #Decision := "FRK_Decisions".EmptyRequest;
   #DecisionAnswer := 0;
   IF #Slot = 0 THEN
       RETURN;
   END_IF;
   IF "FRK_Decisions".Slots[#Slot].RootIndex <> #Owner THEN
       RETURN;
   END_IF;
   #Decision := "FRK_Decisions".Slots[#Slot].Request;
   #DecisionAnswer := "FRK_Decisions".Slots[#Slot].Answer;
END_FUNCTION

FUNCTION "FRK_DecisionRoot" : Int   // FC94, SCL
{ S7_Optimized_Access := 'TRUE' }
VERSION : 0.1
// Core 6.11: one authoritative decision slot per registered root.
// stored: AutoNumber true, IsIECCheckEnabled false, SetENOAutomatically false, UDAEnableTagReadback false
   VAR_INPUT
      Owner : DInt;
      Create : Bool;
   END_VAR
   VAR_TEMP
      RootIndex : DInt;
      Depth : DInt;
      Slot : Int;
   END_VAR
BEGIN

   #FRK_DecisionRoot := 0;
   IF "FRK_Registry".Fault OR "FRK_Registry".Count < 1 OR "FRK_Registry".Count > 32 THEN
       RETURN;
   END_IF;
   #RootIndex := #Owner;
   FOR #Depth := 1 TO 32 DO
       IF #RootIndex < 1 OR #RootIndex > "FRK_Registry".Count THEN
           RETURN;
       END_IF;
       IF NOT "FRK_Registry".Rows[#RootIndex].Valid THEN
           RETURN;
       END_IF;
       IF "FRK_Registry".Rows[#RootIndex].Parent = 0 THEN
           EXIT;
       END_IF;
       #RootIndex := "FRK_Registry".Rows[#RootIndex].Parent;
   END_FOR;
   IF "FRK_Registry".Rows[#RootIndex].Parent <> 0 THEN
       RETURN;
   END_IF;
   FOR #Slot := 1 TO 2 DO
       IF "FRK_Decisions".Slots[#Slot].RootIndex = #RootIndex THEN
           #FRK_DecisionRoot := #Slot;
           RETURN;
       END_IF;
   END_FOR;
   IF NOT #Create THEN
       RETURN;
   END_IF;
   FOR #Slot := 1 TO 2 DO
       IF "FRK_Decisions".Slots[#Slot].RootIndex = 0 THEN
           "FRK_Decisions".Slots[#Slot].RootIndex := #RootIndex;
           #FRK_DecisionRoot := #Slot;
           RETURN;
       END_IF;
   END_FOR;
END_FUNCTION

FUNCTION "FRK_DecisionSubmit" : Bool   // FC98, SCL
{ S7_Optimized_Access := 'TRUE' }
VERSION : 0.1
// stored: AutoNumber true, IsIECCheckEnabled false, SetENOAutomatically false, UDAEnableTagReadback false
   VAR_INPUT
      Owner : DInt;
      OwnerPath : WString;
      Option : DInt;
      Busy : Bool;
      Permit : Bool;
   END_VAR
   VAR_IN_OUT
      Report : "ST_ReleaseReport";
   END_VAR
   VAR_TEMP
      Slot : Int;
      SourcePath : WString[255];
   END_VAR
BEGIN

   #FRK_DecisionSubmit := FALSE;
   #Slot := "FRK_DecisionRoot"(Owner := #Owner, Create := FALSE);
   #SourcePath := #OwnerPath;
   IF NOT #Busy OR #Slot = 0 THEN
       "FRK_ReleaseReason"(Report := #Report,
                           Description := WSTRING#'std.release.noActiveDecision',
                           Reason := 0,
                           Path := #SourcePath,
                           Kind := 4);
       RETURN;
   END_IF;
   IF "FRK_Decisions".Slots[#Slot].RootIndex <> #Owner THEN
       "FRK_ReleaseReason"(Report := #Report,
                           Description := WSTRING#'std.release.noActiveDecision',
                           Reason := 0,
                           Path := #SourcePath,
                           Kind := 4);
       RETURN;
   END_IF;
   IF "FRK_Decisions".Slots[#Slot].Request.Prompt = WSTRING#'' OR "FRK_Decisions".Slots[#Slot].Answer <> 0 THEN
       "FRK_ReleaseReason"(Report := #Report,
                           Description := WSTRING#'std.release.noActiveDecision',
                           Reason := 0,
                           Path := #SourcePath,
                           Kind := 4);
       RETURN;
   END_IF;
   IF #Option < 1 OR #Option > 6 THEN
       "FRK_ReleaseReason"(Report := #Report,
                           Description := WSTRING#'std.release.invalidDecisionOption',
                           Reason := 2008,
                           Path := #SourcePath,
                           Kind := 4);
       RETURN;
   END_IF;
   IF "FRK_Decisions".Slots[#Slot].Request.Options[#Option] = '' THEN
       "FRK_ReleaseReason"(Report := #Report,
                           Description := WSTRING#'std.release.invalidDecisionOption',
                           Reason := 2008,
                           Path := #SourcePath,
                           Kind := 4);
       RETURN;
   END_IF;
   IF NOT #Permit THEN
       "FRK_ReleaseReason"(Report := #Report,
                           Description := WSTRING#'std.release.decisionInterlock',
                           Reason := 2002,
                           Path := #SourcePath,
                           Kind := 3);
       RETURN;
   END_IF;
   IF NOT #Report.Released THEN
       RETURN;
   END_IF;
   "FRK_Decisions".Slots[#Slot].Answer := DINT_TO_INT(#Option);
   #FRK_DecisionSubmit := TRUE;
END_FUNCTION

FUNCTION "FRK_DecisionTake" : Int   // FC100, SCL
{ S7_Optimized_Access := 'TRUE' }
VERSION : 0.1
// stored: AutoNumber true, IsIECCheckEnabled false, SetENOAutomatically false, UDAEnableTagReadback false
   VAR_INPUT
      Owner : DInt;
   END_VAR
   VAR_IN_OUT
      AlarmLog : "FRK_AlarmLog";
   END_VAR
   VAR_TEMP
      Slot : Int;
   END_VAR
BEGIN

   #FRK_DecisionTake := 0;
   #Slot := "FRK_DecisionRoot"(Owner := #Owner, Create := FALSE);
   IF #Slot = 0 THEN
       RETURN;
   END_IF;
   IF "FRK_Decisions".Slots[#Slot].Owner <> #Owner THEN
       RETURN;
   END_IF;
   IF "FRK_Decisions".Slots[#Slot].Answer = 0 THEN
       RETURN;
   END_IF;
   #FRK_DecisionTake := "FRK_Decisions".Slots[#Slot].Answer;
   IF NOT "FRK_Decisions".Slots[#Slot].ResolutionLogged THEN
       "FRK_DecisionAudit"(AlarmLog := #AlarmLog,
                           Key := WSTRING#'std.audit.decisionOperatorResolved',
                           SourcePath := "FRK_Decisions".Slots[#Slot].Request.SourcePath,
                           Option := #FRK_DecisionTake);
   END_IF;
   "FRK_DecisionClear"(Slot := "FRK_Decisions".Slots[#Slot]);
END_FUNCTION

FUNCTION "FRK_DescendantsReady" : Bool   // FC84, SCL
{ S7_Optimized_Access := 'TRUE' }
VERSION : 0.1
// stored: AutoNumber true, IsIECCheckEnabled false, SetENOAutomatically false, UDAEnableTagReadback false
   VAR_INPUT
      OwnerIndex : DInt;
   END_VAR
   VAR_TEMP
      Index : DInt;
      Parent : DInt;
      Depth : DInt;
   END_VAR
BEGIN

   #FRK_DescendantsReady := FALSE;
   IF "FRK_Registry".Fault OR #OwnerIndex < 1 OR #OwnerIndex > "FRK_Registry".Count OR "FRK_Registry".Count > 32 THEN
       RETURN;
   END_IF;
   FOR #Index := 1 TO "FRK_Registry".Count DO
       #Parent := "FRK_Registry".Rows[#Index].Parent;
       FOR #Depth := 1 TO 32 DO
           IF #Parent = #OwnerIndex THEN
               IF "FRK_Registry".Rows[#Index].Exec <> 0 THEN
                   RETURN;
               END_IF;
               EXIT;
           END_IF;
           IF #Parent = 0 THEN
               EXIT;
           END_IF;
           IF #Parent < 1 OR #Parent > "FRK_Registry".Count THEN
               RETURN;
           END_IF;
           #Parent := "FRK_Registry".Rows[#Parent].Parent;
       END_FOR;
       IF #Depth > 32 AND #Parent <> 0 THEN
           RETURN;
       END_IF;
   END_FOR;
   #FRK_DescendantsReady := TRUE;
END_FUNCTION

FUNCTION "FRK_Diagnostic" : Void   // FC8, SCL
{ S7_Optimized_Access := 'TRUE' }
VERSION : 0.1
// stored: AutoNumber true, IsIECCheckEnabled false, SetENOAutomatically false, UDAEnableTagReadback false
   VAR_INPUT
      ReasonCode : DInt;
      Description : WString;
      Severity : DInt;
   END_VAR
   VAR_IN_OUT
      Status : "ST_ModuleStatus";
   END_VAR
   VAR_TEMP
      Stamp : DTL;
      ResultCode : Int;
   END_VAR
BEGIN

   #Status.Diagnostic.ReasonCode := #ReasonCode;
   #Status.Diagnostic.SourcePath := STRING_TO_WSTRING(#Status.Name);
   #Status.Diagnostic.Description := #Description;
   #Status.Diagnostic.IoTag := '';
   #Status.Diagnostic.IoAddress := '';
   #Status.Diagnostic.Severity := #Severity;
   #Status.Diagnostic.Category := 0;
   #ResultCode := RD_SYS_T(OUT => #Stamp);
   IF #ResultCode = 0 THEN
       #Status.Diagnostic.Since := DTL_TO_LDT(#Stamp);
   ELSE
       #Status.Diagnostic.Since := LDT#1970-01-01-00:00:00.000000000;
   END_IF;
   // UTC source alone is not proof of synchronization; quality stays false.
   #Status.Diagnostic.TimeSynchronized := FALSE;
END_FUNCTION

FUNCTION "FRK_Elapsed" : UDInt   // FC5, SCL
{ S7_Optimized_Access := 'TRUE' }
VERSION : 0.1
// stored: AutoNumber true, IsIECCheckEnabled false, SetENOAutomatically false, UDAEnableTagReadback false
   VAR_INPUT
      NewMs : UDInt;
      OldMs : UDInt;
   END_VAR
   VAR_TEMP
      Wide : ULInt;
   END_VAR
BEGIN

   IF #NewMs >= #OldMs THEN
       #Wide := UDINT_TO_ULINT(#NewMs) - UDINT_TO_ULINT(#OldMs);
   ELSE
       #Wide := ULINT#4294967296 + UDINT_TO_ULINT(#NewMs) - UDINT_TO_ULINT(#OldMs);
   END_IF;
   #FRK_Elapsed := ULINT_TO_UDINT(#Wide);
END_FUNCTION

FUNCTION "FRK_End" : Void   // FC19, SCL
{ S7_Optimized_Access := 'TRUE' }
VERSION : 0.1
// stored: AutoNumber true, IsIECCheckEnabled false, SetENOAutomatically false, UDAEnableTagReadback false
   VAR_OUTPUT
      Busy : Bool;
      Done : Bool;
      Error : Bool;
      Aborted : Bool;
      Held : Bool;
      ErrorID : DWord;
      Timing : "ST_ModuleTiming";
   END_VAR
   VAR_IN_OUT
      Core : "FRK_Core";
      Status : "ST_ModuleStatus";
   END_VAR
   VAR_TEMP
      ActiveWide : ULInt;
   END_VAR
BEGIN

   IF #Core.Exec = 1 THEN
       IF #Core.Held AND NOT #Core.HoldReq AND NOT #Core.DiagTouched THEN
           "FRK_ClearDiag"(Status := #Status);
       END_IF;
       // HELD suspends progress timeout. Wall-clock command duration includes it.
       IF NOT #Core.Held AND NOT #Core.HoldReq THEN
           #ActiveWide := UDINT_TO_ULINT(#Core.ActiveMs) + UDINT_TO_ULINT(#Core.DeltaMs);
           IF #ActiveWide > ULINT#2147483647 THEN
               #ActiveWide := ULINT#2147483647;
           END_IF;
           #Core.ActiveMs := ULINT_TO_UDINT(#ActiveWide);
           IF #Core.TimeoutMs > 0 AND #Core.ActiveMs >= #Core.TimeoutMs THEN
               IF #Status.Diagnostic.ReasonCode = 0 THEN
                   "FRK_Fault"(Core := #Core,
                               Status := #Status,
                               ReasonCode := 2001,
                               Description := WSTRING#'fraktal.command.timeout');
               ELSE
                   #Status.Diagnostic.Severity := 1;
                   "FRK_Rationalize"(Diag := #Status.Diagnostic);
                   #Core.Exec := 3;
                   #Core.Step := 0;
                   #Core.Dispatch := FALSE;
               END_IF;
           END_IF;
       END_IF;
   END_IF;
   #Core.Held := #Core.HoldReq AND #Core.Exec = 1;
   IF NOT #Core.Held THEN
       #Core.HoldReason := 0;
   END_IF;
   IF #Core.TimingOpen AND #Core.Exec <> 1 THEN
       "FRK_RecordTiming"(Core := #Core);
   END_IF;
   #Busy := #Core.Exec = 1;
   #Done := #Core.Exec = 2;
   #Error := #Core.Exec = 3;
   #Aborted := #Core.Exec = 4;
   #Held := #Core.Held;
   #ErrorID := DINT_TO_DWORD(#Status.Diagnostic.ReasonCode);
   #Timing := #Core.Timing;
   #Status.State := #Core.Exec;
   #Status.FaultActive := #Core.Exec = 3;
   #Core.HoldReq := FALSE;
   #Core.EvInit := FALSE;
   #Core.EvCommandStart := FALSE;
   #Core.EvAbort := FALSE;
   #Core.EvAbortInError := FALSE;
   #Core.ReleasePending := FALSE;
   "FRK_SyncRegistry"(Index := #Core.RegIndex,
                      Status := #Status);
END_FUNCTION

FUNCTION "FRK_Fault" : Void   // FC9, SCL
{ S7_Optimized_Access := 'TRUE' }
VERSION : 0.1
// stored: AutoNumber true, IsIECCheckEnabled false, SetENOAutomatically false, UDAEnableTagReadback false
   VAR_INPUT
      ReasonCode : DInt;
      Description : WString;
   END_VAR
   VAR_IN_OUT
      Core : "FRK_Core";
      Status : "ST_ModuleStatus";
   END_VAR
BEGIN

   IF #Core.Exec = 3 THEN
       RETURN;
   END_IF;
   "FRK_Diagnostic"(Status := #Status,
                    ReasonCode := #ReasonCode,
                    Description := #Description,
                    Severity := 1);
   "FRK_Rationalize"(Diag := #Status.Diagnostic);
   #Core.Exec := 3;
   #Core.Step := 0;
   #Core.Dispatch := FALSE;
   #Core.DiagTouched := TRUE;
END_FUNCTION

FUNCTION "FRK_Hold" : Void   // FC12, SCL
{ S7_Optimized_Access := 'TRUE' }
VERSION : 0.1
// stored: AutoNumber true, IsIECCheckEnabled false, SetENOAutomatically false, UDAEnableTagReadback false
   VAR_INPUT
      ReasonCode : DInt;
      Description : WString;
   END_VAR
   VAR_IN_OUT
      Core : "FRK_Core";
      Status : "ST_ModuleStatus";
   END_VAR
BEGIN

   IF #Core.Exec <> 1 THEN
       RETURN;
   END_IF;
   IF NOT #Core.Held OR #Core.HoldReason <> #ReasonCode THEN
       "FRK_Diagnostic"(Status := #Status,
                        ReasonCode := #ReasonCode,
                        Description := #Description,
                        Severity := 0);
   END_IF;
   #Core.HoldReq := TRUE;
   #Core.HoldReason := #ReasonCode;
   #Core.DiagTouched := TRUE;
END_FUNCTION

FUNCTION "FRK_HoldDiag" : Void   // FC11, SCL
{ S7_Optimized_Access := 'TRUE' }
VERSION : 0.1
// stored: AutoNumber true, IsIECCheckEnabled false, SetENOAutomatically false, UDAEnableTagReadback false
   VAR_INPUT
      Diag : "ST_Diagnostic";
   END_VAR
   VAR_IN_OUT
      Core : "FRK_Core";
      Status : "ST_ModuleStatus";
   END_VAR
BEGIN

   IF #Core.Exec <> 1 THEN
       RETURN;
   END_IF;
   #Status.Diagnostic := #Diag;
   #Status.Diagnostic.Severity := 0;
   #Core.HoldReq := TRUE;
   #Core.HoldReason := #Diag.ReasonCode;
   #Core.DiagTouched := TRUE;
END_FUNCTION

FUNCTION "FRK_JsonAdd" : Bool   // FC117, SCL
{ S7_Optimized_Access := 'TRUE' }
VERSION : 0.1
// stored: AutoNumber true, IsIECCheckEnabled false, SetENOAutomatically false, UDAEnableTagReadback false
   VAR_INPUT
      Key : String;
      Value : WString;
      Quoted : Bool;
      LastField : Bool;
   END_VAR
   VAR_IN_OUT
      Line : WString;
   END_VAR
   VAR_TEMP
      Index : Int;
      Ch : WChar;
      FirstChar : Int;
      Piece : WString[2];
      Ok : Bool;
   END_VAR
BEGIN

   #FRK_JsonAdd := FALSE;
   #Ok := "FRK_JsonPut"(Text := CONCAT(IN1 := WSTRING#'"', IN2 := STRING_TO_WSTRING(#Key), IN3 := WSTRING#'":'), Line := #Line);
   IF NOT #Ok THEN
       RETURN;
   END_IF;
   IF #Quoted THEN
       #Ok := "FRK_JsonPut"(Text := WSTRING#'"', Line := #Line);
       IF NOT #Ok THEN
           RETURN;
       END_IF;
   END_IF;
   #FirstChar := 1;
   // Siemens integer conversions include a leading '+'. JSON numbers do not.
   IF NOT #Quoted THEN
       IF LEN(#Value) = 0 THEN
           RETURN;
       END_IF;
       IF #Value[1] = WCHAR#'+' THEN
           #FirstChar := 2;
       END_IF;
       IF #FirstChar > LEN(#Value) THEN
           RETURN;
       END_IF;
   END_IF;
   FOR #Index := #FirstChar TO LEN(#Value) DO
       #Ch := #Value[#Index];
       #Piece := WSTRING#' ';
       #Piece[1] := #Ch;
       IF NOT #Quoted AND (#Ch < WCHAR#'0' OR #Ch > WCHAR#'9') THEN
           RETURN;
       END_IF;
       IF #Quoted THEN
           IF #Ch = WCHAR#'"' THEN
               #Piece := WSTRING#'\"';
           ELSIF #Ch = WCHAR#'\' THEN
               #Piece := WSTRING#'\\';
           ELSIF #Ch = WCHAR#'$000A' THEN
               #Piece := WSTRING#'\n';
           ELSIF #Ch = WCHAR#'$000D' THEN
               #Piece := WSTRING#'\r';
           ELSIF #Ch = WCHAR#'$0009' THEN
               #Piece := WSTRING#'\t';
           ELSIF #Ch = WCHAR#'$0008' THEN
               #Piece := WSTRING#'\b';
           ELSIF #Ch = WCHAR#'$000C' THEN
               #Piece := WSTRING#'\f';
           ELSIF #Ch < WCHAR#'$0020' THEN
               RETURN;
           END_IF;
       END_IF;
       #Ok := "FRK_JsonPut"(Text := #Piece, Line := #Line);
       IF NOT #Ok THEN
           RETURN;
       END_IF;
   END_FOR;
   IF #Quoted THEN
       #Ok := "FRK_JsonPut"(Text := WSTRING#'"', Line := #Line);
       IF NOT #Ok THEN
           RETURN;
       END_IF;
   END_IF;
   IF #LastField THEN
       #Piece := WSTRING#'}';
   ELSE
       #Piece := WSTRING#',';
   END_IF;
   #FRK_JsonAdd := "FRK_JsonPut"(Text := #Piece, Line := #Line);
END_FUNCTION

FUNCTION "FRK_JsonHeader" : Bool   // FC126, SCL
{ S7_Optimized_Access := 'TRUE' }
VERSION : 0.1
// stored: AutoNumber true, IsIECCheckEnabled false, SetENOAutomatically false, UDAEnableTagReadback false
   VAR_INPUT
      Data : "ST_ConfigSetInfo";
   END_VAR
   VAR_IN_OUT
      Line : WString;
   END_VAR
   VAR_TEMP
      Ok : Bool;
      Flag : WString[1];
   END_VAR
BEGIN

   #FRK_JsonHeader := FALSE;
   #Line := WSTRING#'{';
   #Ok := "FRK_JsonAdd"(Key := 'set', Value := STRING_TO_WSTRING(#Data.SetName), Quoted := TRUE, LastField := FALSE, Line := #Line);
   IF NOT #Ok THEN
       #Line := WSTRING#'';
       RETURN;
   END_IF;
   #Ok := "FRK_JsonAdd"(Key := 'root', Value := STRING_TO_WSTRING(#Data.RootIdentity), Quoted := TRUE, LastField := FALSE, Line := #Line);
   IF NOT #Ok THEN
       #Line := WSTRING#'';
       RETURN;
   END_IF;
   #Ok := "FRK_JsonAdd"(Key := 'schema', Value := UINT_TO_WSTRING(#Data.SetSchema), Quoted := FALSE, LastField := FALSE, Line := #Line);
   IF NOT #Ok THEN
       #Line := WSTRING#'';
       RETURN;
   END_IF;
   #Ok := "FRK_JsonAdd"(Key := 'configRev', Value := UDINT_TO_WSTRING(#Data.ConfigRev), Quoted := FALSE, LastField := FALSE, Line := #Line);
   IF NOT #Ok THEN
       #Line := WSTRING#'';
       RETURN;
   END_IF;
   #Ok := "FRK_JsonAdd"(Key := 'kind', Value := DINT_TO_WSTRING(#Data.Kind), Quoted := FALSE, LastField := FALSE, Line := #Line);
   IF NOT #Ok THEN
       #Line := WSTRING#'';
       RETURN;
   END_IF;
   #Ok := "FRK_JsonAdd"(Key := 'model', Value := STRING_TO_WSTRING(#Data.ModelCode), Quoted := TRUE, LastField := FALSE, Line := #Line);
   IF NOT #Ok THEN
       #Line := WSTRING#'';
       RETURN;
   END_IF;
   #Ok := "FRK_JsonAdd"(Key := 'records', Value := DINT_TO_WSTRING(#Data.RecordCount), Quoted := FALSE, LastField := FALSE, Line := #Line);
   IF NOT #Ok THEN
       #Line := WSTRING#'';
       RETURN;
   END_IF;
   #Ok := "FRK_JsonAdd"(Key := 'created', Value := ULINT_TO_WSTRING(LDT_TO_ULINT(#Data.CreatedAt) / ULINT#1000000000), Quoted := FALSE, LastField := FALSE, Line := #Line);
   IF NOT #Ok THEN
       #Line := WSTRING#'';
       RETURN;
   END_IF;
   IF #Data.TimeSynchronized THEN
       #Flag := WSTRING#'1';
   ELSE
       #Flag := WSTRING#'0';
   END_IF;
   #Ok := "FRK_JsonAdd"(Key := 'clock', Value := #Flag, Quoted := FALSE, LastField := TRUE, Line := #Line);
   IF NOT #Ok THEN
       #Line := WSTRING#'';
       RETURN;
   END_IF;
   #FRK_JsonHeader := TRUE;
END_FUNCTION

FUNCTION "FRK_JsonParse" : Bool   // FC118, SCL
{ S7_Optimized_Access := 'TRUE' }
VERSION : 0.1
// Strict flat JSON object scanner: whole object, unique known fields, exact
//  types, numeric integer grammar; strings decode escapes before owner checks.
// stored: AutoNumber true, IsIECCheckEnabled false, SetENOAutomatically false, UDAEnableTagReadback false
   VAR_INPUT
      Line : WString;
   END_VAR
   VAR_IN_OUT
      Fields : Array[1..9] of "FRK_JsonField";
      Count : Int;
   END_VAR
   VAR_TEMP
      Pos : Int;
      Limit : Int;
      Digit : Int;
      CodePoint : UInt;
      HexIndex : Int;
      Index : Int;
      Part : Int;
      Text : WString[160];
      Piece : WString[1];
      Quoted : Bool;
      Closed : Bool;
      Ch : WChar;
   END_VAR
BEGIN

   #FRK_JsonParse := FALSE;
   #Count := 0;
   #Pos := 1;
   #Limit := LEN(#Line);
   IF #Limit < 2 OR #Line[#Pos] <> WCHAR#'{' THEN
       RETURN;
   END_IF;
   #Pos := #Pos + 1;
   WHILE #Pos <= #Limit DO
       "FRK_JsonSkip"(Line := #Line,
                      Pos := #Pos);
       IF #Pos > #Limit OR #Count >= 9 THEN
           RETURN;
       END_IF;
       #Count := #Count + 1;
       FOR #Part := 1 TO 2 DO
           #Text := WSTRING#'';
           #Closed := FALSE;
           #Quoted := #Line[#Pos] = WCHAR#'"';
           IF #Part = 1 AND NOT #Quoted THEN
               RETURN;
           END_IF;
           IF #Quoted THEN
               #Pos := #Pos + 1;
           END_IF;
           WHILE #Pos <= #Limit DO
               #Ch := #Line[#Pos];
               IF #Quoted AND #Ch = WCHAR#'"' THEN
                   #Closed := TRUE;
                   #Pos := #Pos + 1;
                   EXIT;
               END_IF;
               IF NOT #Quoted AND (#Ch = WCHAR#',' OR #Ch = WCHAR#'}' OR #Ch = WCHAR#' ') THEN
                   #Closed := TRUE;
                   EXIT;
               END_IF;
               IF #Ch < WCHAR#'$0020' THEN
                   RETURN;
               END_IF;
               IF #Quoted AND #Ch = WCHAR#'\' THEN
                   #Pos := #Pos + 1;
                   IF #Pos > #Limit THEN
                       RETURN;
                   END_IF;
                   #Ch := #Line[#Pos];
                   IF #Ch = WCHAR#'u' THEN
                       #CodePoint := 0;
                       FOR #HexIndex := 1 TO 4 DO
                           #Pos := #Pos + 1;
                           IF #Pos > #Limit THEN
                               RETURN;
                           END_IF;
                           #Ch := #Line[#Pos];
                           #Digit := -1;
                           IF #Ch >= WCHAR#'0' AND #Ch <= WCHAR#'9' THEN
                               #Digit := WORD_TO_INT(WCHAR_TO_WORD(#Ch)) - 48;
                           ELSIF #Ch >= WCHAR#'a' AND #Ch <= WCHAR#'f' THEN
                               #Digit := WORD_TO_INT(WCHAR_TO_WORD(#Ch)) - 87;
                           ELSIF #Ch >= WCHAR#'A' AND #Ch <= WCHAR#'F' THEN
                               #Digit := WORD_TO_INT(WCHAR_TO_WORD(#Ch)) - 55;
                           END_IF;
                           IF #Digit < 0 THEN
                               RETURN;
                           END_IF;
                           #CodePoint := #CodePoint * 16 + INT_TO_UINT(#Digit);
                       END_FOR;
                       IF #CodePoint = 0 OR #CodePoint >= UINT#16#D000 THEN
                           RETURN;
                       END_IF;
                       #Ch := WORD_TO_WCHAR(UINT_TO_WORD(#CodePoint));
                   ELSIF #Ch = WCHAR#'n' THEN
                       #Ch := WCHAR#'$000A';
                   ELSIF #Ch = WCHAR#'r' THEN
                       #Ch := WCHAR#'$000D';
                   ELSIF #Ch = WCHAR#'t' THEN
                       #Ch := WCHAR#'$0009';
                   ELSIF #Ch = WCHAR#'b' THEN
                       #Ch := WCHAR#'$0008';
                   ELSIF #Ch = WCHAR#'f' THEN
                       #Ch := WCHAR#'$000C';
                   ELSIF #Ch <> WCHAR#'"' AND #Ch <> WCHAR#'\' AND #Ch <> WCHAR#'/' THEN
                       RETURN;
                   END_IF;
               ELSIF NOT #Quoted AND (#Ch < WCHAR#'0' OR #Ch > WCHAR#'9') THEN
                   RETURN;
               END_IF;
               IF LEN(#Text) >= 160 THEN
                   RETURN;
               END_IF;
               #Piece := WSTRING#' ';
               #Piece[1] := #Ch;
               #Text := CONCAT(IN1 := #Text, IN2 := #Piece);
               #Pos := #Pos + 1;
           END_WHILE;
           IF NOT #Closed THEN
               RETURN;
           END_IF;
           IF #Part = 1 THEN
               IF LEN(#Text) < 1 OR LEN(#Text) > 16 THEN
                   RETURN;
               END_IF;
               #Fields[#Count].Key := WSTRING_TO_STRING(#Text);
               FOR #Index := 1 TO #Count - 1 DO
                   IF #Fields[#Index].Key = #Fields[#Count].Key THEN
                       RETURN;
                   END_IF;
               END_FOR;
               "FRK_JsonSkip"(Line := #Line,
                              Pos := #Pos);
               IF #Pos > #Limit THEN
                   RETURN;
               END_IF;
               IF #Line[#Pos] <> WCHAR#':' THEN
                   RETURN;
               END_IF;
               #Pos := #Pos + 1;
               "FRK_JsonSkip"(Line := #Line,
                              Pos := #Pos);
               IF #Pos > #Limit THEN
                   RETURN;
               END_IF;
           ELSE
               IF NOT #Quoted AND (LEN(#Text) = 0 OR (LEN(#Text) > 1 AND #Text[1] = WCHAR#'0')) THEN
                   RETURN;
               END_IF;
               #Fields[#Count].Text := #Text;
               #Fields[#Count].Quoted := #Quoted;
           END_IF;
       END_FOR;
       "FRK_JsonSkip"(Line := #Line,
                      Pos := #Pos);
       IF #Pos > #Limit THEN
           RETURN;
       END_IF;
       IF #Line[#Pos] = WCHAR#'}' THEN
           #Pos := #Pos + 1;
           "FRK_JsonSkip"(Line := #Line,
                          Pos := #Pos);
           #FRK_JsonParse := #Pos > #Limit;
           RETURN;
       END_IF;
       IF #Line[#Pos] <> WCHAR#',' THEN
           RETURN;
       END_IF;
       #Pos := #Pos + 1;
   END_WHILE;
END_FUNCTION

FUNCTION "FRK_JsonPut" : Bool   // FC116, SCL
{ S7_Optimized_Access := 'TRUE' }
VERSION : 0.1
// Append complete text or refuse. Explicit destination width and length check
//  protect long WSTRING lines against truncation in the Siemens string runtime.
// stored: AutoNumber true, IsIECCheckEnabled false, SetENOAutomatically false, UDAEnableTagReadback false
   VAR_INPUT
      Text : WString;
   END_VAR
   VAR_IN_OUT
      Line : WString;
   END_VAR
   VAR_TEMP
      Expected : Int;
   END_VAR
BEGIN

   #FRK_JsonPut := FALSE;
   #Expected := LEN(#Line) + LEN(#Text);
   IF #Expected > 480 THEN
       RETURN;
   END_IF;
   #Line := CONCAT(IN1 := #Line, IN2 := #Text);
   #FRK_JsonPut := LEN(#Line) = #Expected;
END_FUNCTION

FUNCTION "FRK_JsonReadHeader" : Bool   // FC127, SCL
{ S7_Optimized_Access := 'TRUE' }
VERSION : 0.1
// stored: AutoNumber true, IsIECCheckEnabled false, SetENOAutomatically false, UDAEnableTagReadback false
   VAR_INPUT
      Count : Int;
      Fields : Array[1..9] of "FRK_JsonField";
   END_VAR
   VAR_IN_OUT
      Data : "ST_ConfigSetInfo";
   END_VAR
   VAR_TEMP
      Candidate : "ST_ConfigSetInfo";
      Index : Int;
      Found : Int;
      Ok : Bool;
   END_VAR
BEGIN

   #FRK_JsonReadHeader := FALSE;
   IF #Count <> 9 THEN
       RETURN;
   END_IF;
   #Found := 0;
   FOR #Index := 1 TO #Count DO
       IF #Fields[#Index].Key = 'set' THEN
           #Found := #Index;
       END_IF;
   END_FOR;
   IF #Found = 0 THEN
       RETURN;
   END_IF;
   IF #Fields[#Found].Quoted <> TRUE THEN
       RETURN;
   END_IF;
   IF LEN(#Fields[#Found].Text) > 80 OR STRING_TO_WSTRING(WSTRING_TO_STRING(#Fields[#Found].Text)) <> #Fields[#Found].Text THEN
       RETURN;
   END_IF;
   #Candidate.SetName := WSTRING_TO_STRING(#Fields[#Found].Text);
   #Found := 0;
   FOR #Index := 1 TO #Count DO
       IF #Fields[#Index].Key = 'root' THEN
           #Found := #Index;
       END_IF;
   END_FOR;
   IF #Found = 0 THEN
       RETURN;
   END_IF;
   IF #Fields[#Found].Quoted <> TRUE THEN
       RETURN;
   END_IF;
   IF LEN(#Fields[#Found].Text) > 80 OR STRING_TO_WSTRING(WSTRING_TO_STRING(#Fields[#Found].Text)) <> #Fields[#Found].Text THEN
       RETURN;
   END_IF;
   #Candidate.RootIdentity := WSTRING_TO_STRING(#Fields[#Found].Text);
   #Found := 0;
   FOR #Index := 1 TO #Count DO
       IF #Fields[#Index].Key = 'schema' THEN
           #Found := #Index;
       END_IF;
   END_FOR;
   IF #Found = 0 THEN
       RETURN;
   END_IF;
   IF #Fields[#Found].Quoted <> FALSE THEN
       RETURN;
   END_IF;
   #Ok := "FRK_ConfigDecode"(Text := #Fields[#Found].Text, Storage := 4, Minimum := 0.0, Maximum := 65535.0, MaxLength := 0, Value := "FRK_ConfigScratch".Value);
   IF NOT #Ok THEN
       RETURN;
   END_IF;
   #Candidate.SetSchema := LINT_TO_UINT("FRK_ConfigScratch".Value.Number);
   #Found := 0;
   FOR #Index := 1 TO #Count DO
       IF #Fields[#Index].Key = 'configRev' THEN
           #Found := #Index;
       END_IF;
   END_FOR;
   IF #Found = 0 THEN
       RETURN;
   END_IF;
   IF #Fields[#Found].Quoted <> FALSE THEN
       RETURN;
   END_IF;
   #Ok := "FRK_ConfigDecode"(Text := #Fields[#Found].Text, Storage := 4, Minimum := 0.0, Maximum := 4294967295.0, MaxLength := 0, Value := "FRK_ConfigScratch".Value);
   IF NOT #Ok THEN
       RETURN;
   END_IF;
   #Candidate.ConfigRev := LINT_TO_UDINT("FRK_ConfigScratch".Value.Number);
   #Found := 0;
   FOR #Index := 1 TO #Count DO
       IF #Fields[#Index].Key = 'kind' THEN
           #Found := #Index;
       END_IF;
   END_FOR;
   IF #Found = 0 THEN
       RETURN;
   END_IF;
   IF #Fields[#Found].Quoted <> FALSE THEN
       RETURN;
   END_IF;
   #Ok := "FRK_ConfigDecode"(Text := #Fields[#Found].Text, Storage := 4, Minimum := 0.0, Maximum := 1.0, MaxLength := 0, Value := "FRK_ConfigScratch".Value);
   IF NOT #Ok THEN
       RETURN;
   END_IF;
   #Candidate.Kind := LINT_TO_DINT("FRK_ConfigScratch".Value.Number);
   #Found := 0;
   FOR #Index := 1 TO #Count DO
       IF #Fields[#Index].Key = 'model' THEN
           #Found := #Index;
       END_IF;
   END_FOR;
   IF #Found = 0 THEN
       RETURN;
   END_IF;
   IF #Fields[#Found].Quoted <> TRUE THEN
       RETURN;
   END_IF;
   IF LEN(#Fields[#Found].Text) > 64 OR STRING_TO_WSTRING(WSTRING_TO_STRING(#Fields[#Found].Text)) <> #Fields[#Found].Text THEN
       RETURN;
   END_IF;
   #Candidate.ModelCode := WSTRING_TO_STRING(#Fields[#Found].Text);
   #Found := 0;
   FOR #Index := 1 TO #Count DO
       IF #Fields[#Index].Key = 'records' THEN
           #Found := #Index;
       END_IF;
   END_FOR;
   IF #Found = 0 THEN
       RETURN;
   END_IF;
   IF #Fields[#Found].Quoted <> FALSE THEN
       RETURN;
   END_IF;
   #Ok := "FRK_ConfigDecode"(Text := #Fields[#Found].Text, Storage := 4, Minimum := 0.0, Maximum := 24.0, MaxLength := 0, Value := "FRK_ConfigScratch".Value);
   IF NOT #Ok THEN
       RETURN;
   END_IF;
   #Candidate.RecordCount := LINT_TO_INT("FRK_ConfigScratch".Value.Number);
   #Found := 0;
   FOR #Index := 1 TO #Count DO
       IF #Fields[#Index].Key = 'created' THEN
           #Found := #Index;
       END_IF;
   END_FOR;
   IF #Found = 0 THEN
       RETURN;
   END_IF;
   IF #Fields[#Found].Quoted <> FALSE THEN
       RETURN;
   END_IF;
   #Ok := "FRK_ConfigDecode"(Text := #Fields[#Found].Text, Storage := 4, Minimum := 0.0, Maximum := 4294967295.0, MaxLength := 0, Value := "FRK_ConfigScratch".Value);
   IF NOT #Ok THEN
       RETURN;
   END_IF;
   #Candidate.CreatedAt := ULINT_TO_LDT(LINT_TO_ULINT("FRK_ConfigScratch".Value.Number) * ULINT#1000000000);
   #Found := 0;
   FOR #Index := 1 TO #Count DO
       IF #Fields[#Index].Key = 'clock' THEN
           #Found := #Index;
       END_IF;
   END_FOR;
   IF #Found = 0 THEN
       RETURN;
   END_IF;
   IF #Fields[#Found].Quoted <> FALSE THEN
       RETURN;
   END_IF;
   #Ok := "FRK_ConfigDecode"(Text := #Fields[#Found].Text, Storage := 4, Minimum := 0.0, Maximum := 1.0, MaxLength := 0, Value := "FRK_ConfigScratch".Value);
   IF NOT #Ok THEN
       RETURN;
   END_IF;
   #Candidate.TimeSynchronized := "FRK_ConfigScratch".Value.Number = 1;
   #Data := #Candidate;
   #FRK_JsonReadHeader := TRUE;
END_FUNCTION

FUNCTION "FRK_JsonReadRecord" : Bool   // FC129, SCL
{ S7_Optimized_Access := 'TRUE' }
VERSION : 0.1
// stored: AutoNumber true, IsIECCheckEnabled false, SetENOAutomatically false, UDAEnableTagReadback false
   VAR_INPUT
      Count : Int;
      Fields : Array[1..9] of "FRK_JsonField";
   END_VAR
   VAR_IN_OUT
      Data : "ST_ConfigRecord";
   END_VAR
   VAR_TEMP
      Candidate : "ST_ConfigRecord";
      Index : Int;
      Found : Int;
      Ok : Bool;
   END_VAR
BEGIN

   #FRK_JsonReadRecord := FALSE;
   IF #Count <> 6 THEN
       RETURN;
   END_IF;
   #Found := 0;
   FOR #Index := 1 TO #Count DO
       IF #Fields[#Index].Key = 'scope' THEN
           #Found := #Index;
       END_IF;
   END_FOR;
   IF #Found = 0 THEN
       RETURN;
   END_IF;
   IF #Fields[#Found].Quoted <> TRUE THEN
       RETURN;
   END_IF;
   IF LEN(#Fields[#Found].Text) > 80 OR STRING_TO_WSTRING(WSTRING_TO_STRING(#Fields[#Found].Text)) <> #Fields[#Found].Text THEN
       RETURN;
   END_IF;
   #Candidate.Scope := WSTRING_TO_STRING(#Fields[#Found].Text);
   #Found := 0;
   FOR #Index := 1 TO #Count DO
       IF #Fields[#Index].Key = 'key' THEN
           #Found := #Index;
       END_IF;
   END_FOR;
   IF #Found = 0 THEN
       RETURN;
   END_IF;
   IF #Fields[#Found].Quoted <> TRUE THEN
       RETURN;
   END_IF;
   IF LEN(#Fields[#Found].Text) > 160 OR STRING_TO_WSTRING(WSTRING_TO_STRING(#Fields[#Found].Text)) <> #Fields[#Found].Text THEN
       RETURN;
   END_IF;
   #Candidate.WriteKey := WSTRING_TO_STRING(#Fields[#Found].Text);
   #Found := 0;
   FOR #Index := 1 TO #Count DO
       IF #Fields[#Index].Key = 'rev' THEN
           #Found := #Index;
       END_IF;
   END_FOR;
   IF #Found = 0 THEN
       RETURN;
   END_IF;
   IF #Fields[#Found].Quoted <> FALSE THEN
       RETURN;
   END_IF;
   #Ok := "FRK_ConfigDecode"(Text := #Fields[#Found].Text, Storage := 4, Minimum := 0.0, Maximum := 4294967295.0, MaxLength := 0, Value := "FRK_ConfigScratch".Value);
   IF NOT #Ok THEN
       RETURN;
   END_IF;
   #Candidate.Revision := LINT_TO_UDINT("FRK_ConfigScratch".Value.Number);
   #Found := 0;
   FOR #Index := 1 TO #Count DO
       IF #Fields[#Index].Key = 'kind' THEN
           #Found := #Index;
       END_IF;
   END_FOR;
   IF #Found = 0 THEN
       RETURN;
   END_IF;
   IF #Fields[#Found].Quoted <> FALSE THEN
       RETURN;
   END_IF;
   #Ok := "FRK_ConfigDecode"(Text := #Fields[#Found].Text, Storage := 4, Minimum := 0.0, Maximum := 1.0, MaxLength := 0, Value := "FRK_ConfigScratch".Value);
   IF NOT #Ok THEN
       RETURN;
   END_IF;
   #Candidate.Kind := LINT_TO_DINT("FRK_ConfigScratch".Value.Number);
   #Found := 0;
   FOR #Index := 1 TO #Count DO
       IF #Fields[#Index].Key = 'type' THEN
           #Found := #Index;
       END_IF;
   END_FOR;
   IF #Found = 0 THEN
       RETURN;
   END_IF;
   IF #Fields[#Found].Quoted <> FALSE THEN
       RETURN;
   END_IF;
   #Ok := "FRK_ConfigDecode"(Text := #Fields[#Found].Text, Storage := 4, Minimum := 0.0, Maximum := 3.0, MaxLength := 0, Value := "FRK_ConfigScratch".Value);
   IF NOT #Ok THEN
       RETURN;
   END_IF;
   #Candidate.ValueType := LINT_TO_DINT("FRK_ConfigScratch".Value.Number);
   #Found := 0;
   FOR #Index := 1 TO #Count DO
       IF #Fields[#Index].Key = 'value' THEN
           #Found := #Index;
       END_IF;
   END_FOR;
   IF #Found = 0 THEN
       RETURN;
   END_IF;
   IF #Fields[#Found].Quoted <> TRUE THEN
       RETURN;
   END_IF;
   IF LEN(#Fields[#Found].Text) > 80 OR STRING_TO_WSTRING(WSTRING_TO_STRING(#Fields[#Found].Text)) <> #Fields[#Found].Text THEN
       RETURN;
   END_IF;
   #Candidate.ValueText := WSTRING_TO_STRING(#Fields[#Found].Text);
   #Data := #Candidate;
   #FRK_JsonReadRecord := TRUE;
END_FUNCTION

FUNCTION "FRK_JsonRecord" : Bool   // FC128, SCL
{ S7_Optimized_Access := 'TRUE' }
VERSION : 0.1
// stored: AutoNumber true, IsIECCheckEnabled false, SetENOAutomatically false, UDAEnableTagReadback false
   VAR_INPUT
      Data : "ST_ConfigRecord";
   END_VAR
   VAR_IN_OUT
      Line : WString;
   END_VAR
   VAR_TEMP
      Ok : Bool;
      Flag : WString[1];
   END_VAR
BEGIN

   #FRK_JsonRecord := FALSE;
   #Line := WSTRING#'{';
   #Ok := "FRK_JsonAdd"(Key := 'scope', Value := STRING_TO_WSTRING(#Data.Scope), Quoted := TRUE, LastField := FALSE, Line := #Line);
   IF NOT #Ok THEN
       #Line := WSTRING#'';
       RETURN;
   END_IF;
   #Ok := "FRK_JsonAdd"(Key := 'key', Value := STRING_TO_WSTRING(#Data.WriteKey), Quoted := TRUE, LastField := FALSE, Line := #Line);
   IF NOT #Ok THEN
       #Line := WSTRING#'';
       RETURN;
   END_IF;
   #Ok := "FRK_JsonAdd"(Key := 'rev', Value := UDINT_TO_WSTRING(#Data.Revision), Quoted := FALSE, LastField := FALSE, Line := #Line);
   IF NOT #Ok THEN
       #Line := WSTRING#'';
       RETURN;
   END_IF;
   #Ok := "FRK_JsonAdd"(Key := 'kind', Value := DINT_TO_WSTRING(#Data.Kind), Quoted := FALSE, LastField := FALSE, Line := #Line);
   IF NOT #Ok THEN
       #Line := WSTRING#'';
       RETURN;
   END_IF;
   #Ok := "FRK_JsonAdd"(Key := 'type', Value := DINT_TO_WSTRING(#Data.ValueType), Quoted := FALSE, LastField := FALSE, Line := #Line);
   IF NOT #Ok THEN
       #Line := WSTRING#'';
       RETURN;
   END_IF;
   #Ok := "FRK_JsonAdd"(Key := 'value', Value := STRING_TO_WSTRING(#Data.ValueText), Quoted := TRUE, LastField := TRUE, Line := #Line);
   IF NOT #Ok THEN
       #Line := WSTRING#'';
       RETURN;
   END_IF;
   #FRK_JsonRecord := TRUE;
END_FUNCTION

FUNCTION "FRK_JsonSkip" : Void   // FC121, SCL
{ S7_Optimized_Access := 'TRUE' }
VERSION : 0.1
// stored: AutoNumber true, IsIECCheckEnabled false, SetENOAutomatically false, UDAEnableTagReadback false
   VAR_INPUT
      Line : WString;
   END_VAR
   VAR_IN_OUT
      Pos : Int;
   END_VAR
BEGIN

   WHILE #Pos <= LEN(#Line) DO
       IF #Line[#Pos] <> WCHAR#' ' AND #Line[#Pos] <> WCHAR#'$0009' AND #Line[#Pos] <> WCHAR#'$000A' AND #Line[#Pos] <> WCHAR#'$000D' THEN
           RETURN;
       END_IF;
       #Pos := #Pos + 1;
   END_WHILE;
END_FUNCTION

FUNCTION "FRK_ManualApply" : Void   // FC90, SCL
{ S7_Optimized_Access := 'TRUE' }
VERSION : 0.1
// stored: AutoNumber true, IsIECCheckEnabled false, SetENOAutomatically false, UDAEnableTagReadback false
   VAR_INPUT
      Request : "ST_HmiRequest";
      Status : "ST_ModuleStatus";
      Core : "FRK_Core";
      Commands : Array[1..12] of "ST_CommandInfo";
      Count : DInt;
      Conditions : Array[1..16] of "FRK_ManualConditionRow";
   END_VAR
   VAR_IN_OUT
      Report : "ST_ReleaseReport";
      Execute : Bool;
      Command : DInt;
      ManualOwned : Bool;
   END_VAR
   VAR_TEMP
      Index : Int;
      Supported : Bool;
      PreviousCount : Int;
   END_VAR
BEGIN

   #Supported := FALSE;
   IF #Count >= 0 AND #Count <= 12 THEN
       FOR #Index := 1 TO DINT_TO_INT(#Count) DO
           IF #Commands[#Index].Value = #Request.IntValue AND #Commands[#Index].Style = 0 THEN
               #Supported := TRUE;
           END_IF;
       END_FOR;
   END_IF;
   IF NOT #Supported THEN
       "FRK_ReleaseReason"(Report := #Report,
                           Description := WSTRING#'std.error.unsupportedHmiRequest',
                           Reason := 2008,
                           Path := STRING_TO_WSTRING(#Status.Name),
                           Kind := 4);
   END_IF;
   IF #Core.Exec <> 0 OR #Execute OR #Core.ReleasePending THEN
       "FRK_ReleaseReason"(Report := #Report,
                           Description := WSTRING#'std.error.hmiRequestRejected',
                           Reason := 2011,
                           Path := STRING_TO_WSTRING(#Status.Name),
                           Kind := 4);
   END_IF;
   FOR #Index := 1 TO 16 DO
       IF #Conditions[#Index].Used AND NOT #Conditions[#Index].Ok THEN
           IF #Conditions[#Index].Value = 0 OR #Conditions[#Index].Value = #Request.IntValue THEN
               #PreviousCount := #Report.Count;
               "FRK_ReleaseReason"(Report := #Report,
                                   Description := #Conditions[#Index].Diag.Description,
                                   Reason := #Conditions[#Index].Diag.ReasonCode,
                                   Path := STRING_TO_WSTRING(#Status.Name),
                                   Kind := 3);
               IF #Report.Count > #PreviousCount THEN
                   #Report.Reasons[#Report.Count].Bypassable := #Conditions[#Index].Bypassable;
               END_IF;
           END_IF;
       END_IF;
   END_FOR;
   IF #Request.Kind = 11 AND #Report.Released THEN
       #Command := #Request.IntValue;
       #Execute := TRUE;
       #ManualOwned := TRUE;
   END_IF;
END_FUNCTION

FUNCTION "FRK_ManualCommon" : Void   // FC88, SCL
{ S7_Optimized_Access := 'TRUE' }
VERSION : 0.1
// stored: AutoNumber true, IsIECCheckEnabled false, SetENOAutomatically false, UDAEnableTagReadback false
   VAR_INPUT
      Core : "FRK_Core";
      Unit : "FRK_Unit";
      Status : "ST_ModuleStatus";
   END_VAR
   VAR_IN_OUT
      Report : "ST_ReleaseReport";
   END_VAR
BEGIN

   IF #Unit.Mode <> 1 OR #Unit.ModePending THEN
       "FRK_ReleaseReason"(Report := #Report,
                           Description := WSTRING#'std.release.manualModeRequired',
                           Reason := 2002,
                           Path := STRING_TO_WSTRING(#Status.Name),
                           Kind := 0);
   END_IF;
   IF #Core.Exec <> 0 OR #Unit.Clearing OR #Unit.FaultLatched THEN
       "FRK_ReleaseReason"(Report := #Report,
                           Description := WSTRING#'std.error.hmiRequestRejected',
                           Reason := 2011,
                           Path := STRING_TO_WSTRING(#Status.Name),
                           Kind := 4);
   END_IF;
   IF #Unit.AlarmBlocking THEN
       "FRK_ReleaseReason"(Report := #Report,
                           Description := WSTRING#'std.release.manualReset',
                           Reason := 0,
                           Path := STRING_TO_WSTRING(#Status.Name),
                           Kind := 2);
   END_IF;
   IF NOT #Unit.Permit THEN
       "FRK_ReleaseReason"(Report := #Report,
                           Description := #Unit.PermitDiag.Description,
                           Reason := #Unit.PermitDiag.ReasonCode,
                           Path := #Unit.PermitDiag.SourcePath,
                           Kind := 3);
   END_IF;
END_FUNCTION

FUNCTION "FRK_ManualCondition" : Void   // FC89, SCL
{ S7_Optimized_Access := 'TRUE' }
VERSION : 0.1
// stored: AutoNumber true, IsIECCheckEnabled false, SetENOAutomatically false, UDAEnableTagReadback false
   VAR_INPUT
      Slot : Int;
      Value : DInt;
      Ok : Bool;
      Diag : "ST_Diagnostic";
      Bypassable : Bool;
   END_VAR
   VAR_IN_OUT
      Conditions : Array[1..16] of "FRK_ManualConditionRow";
   END_VAR
BEGIN

   IF #Slot < 1 OR #Slot > 16 THEN
       RETURN;
   END_IF;
   #Conditions[#Slot].Used := TRUE;
   #Conditions[#Slot].Value := #Value;
   #Conditions[#Slot].Ok := #Ok;
   #Conditions[#Slot].Diag := #Diag;
   #Conditions[#Slot].Bypassable := #Bypassable;
END_FUNCTION

FUNCTION "FRK_ManualFinish" : Void   // FC91, SCL
{ S7_Optimized_Access := 'TRUE' }
VERSION : 0.1
// stored: AutoNumber true, IsIECCheckEnabled false, SetENOAutomatically false, UDAEnableTagReadback false
   VAR_INPUT
      Core : "FRK_Core";
   END_VAR
   VAR_IN_OUT
      Execute : Bool;
      ManualOwned : Bool;
   END_VAR
BEGIN

   IF #ManualOwned AND #Core.Exec <> 1 THEN
       #Execute := FALSE;
       #ManualOwned := FALSE;
   END_IF;
END_FUNCTION

FUNCTION "FRK_PartAborted" : Void   // FC75, SCL
{ S7_Optimized_Access := 'TRUE' }
VERSION : 0.1
// stored: AutoNumber true, IsIECCheckEnabled false, SetENOAutomatically false, UDAEnableTagReadback false
   VAR_IN_OUT
      Core : "FRK_Core";
      Unit : "FRK_Unit";
      Status : "ST_ModuleStatus";
      Part : "ST_PartContext";
      AlarmLog : "FRK_AlarmLog";
   END_VAR
BEGIN

   IF #Unit.CarrierIndex = 0 OR NOT #Part.Present THEN
       RETURN;
   END_IF;
   #Part.Result.Verdict := 0;
   IF #Core.Exec = 3 AND #Part.Result.ReasonCode = 0 THEN
       #Part.Result.ReasonCode := #Status.Diagnostic.ReasonCode;
   END_IF;
   "FRK_PartEvent"(AlarmLog := #AlarmLog,
                   Reason := 2027,
                   Uid := #Part.Uid,
                   SourcePath := #Status.Name);
   #Part.Present := FALSE;
END_FUNCTION

FUNCTION "FRK_PartEvent" : Void   // FC71, SCL
{ S7_Optimized_Access := 'TRUE' }
VERSION : 0.1
// stored: AutoNumber true, IsIECCheckEnabled false, SetENOAutomatically false, UDAEnableTagReadback false
   VAR_INPUT
      Reason : DInt;
      Uid : String;
      SourcePath : String;
   END_VAR
   VAR_IN_OUT
      AlarmLog : "FRK_AlarmLog";
   END_VAR
   VAR_TEMP
      Description : WString[255];
   END_VAR
BEGIN

   CASE #Reason OF
       2024:
           #Description := WSTRING#'std.event.partReceived: ';
       2025:
           #Description := WSTRING#'std.event.partProcessingStarted: ';
       2026:
           #Description := WSTRING#'std.event.partProcessed: ';
       2027:
           #Description := WSTRING#'std.event.partAborted: ';
       ELSE
           #Description := WSTRING#'';
   END_CASE;
   #Description := CONCAT(IN1 := #Description, IN2 := STRING_TO_WSTRING(#Uid));
   "FRK_AlarmMessage"(AlarmLog := #AlarmLog,
                      Reason := #Reason,
                      Description := #Description,
                      SourcePath := STRING_TO_WSTRING(#SourcePath));
END_FUNCTION

FUNCTION "FRK_PartProcessed" : Bool   // FC74, SCL
{ S7_Optimized_Access := 'TRUE' }
VERSION : 0.1
// stored: AutoNumber true, IsIECCheckEnabled false, SetENOAutomatically false, UDAEnableTagReadback false
   VAR_INPUT
      Verdict : DInt;
      Reason : DInt;
   END_VAR
   VAR_IN_OUT
      Core : "FRK_Core";
      Unit : "FRK_Unit";
      Status : "ST_ModuleStatus";
      Part : "ST_PartContext";
      AlarmLog : "FRK_AlarmLog";
   END_VAR
   VAR_TEMP
      Index : DInt;
      Stamp : DTL;
      ResultCode : Int;
   END_VAR
BEGIN

   #FRK_PartProcessed := FALSE;
   #Index := #Unit.CarrierIndex;
   IF #Index = 0 OR NOT #Part.Present THEN
       RETURN;
   END_IF;
   IF #Verdict < 1 OR #Verdict > 3 OR (#Verdict = 2 AND #Reason = 0) THEN
       "FRK_Fault"(Core := #Core,
                   Status := #Status,
                   ReasonCode := 2023,
                   Description := WSTRING#'std.error.nokReasonRequired');
       RETURN;
   END_IF;
   IF #Index < 1 OR #Index > 32 THEN
       "FRK_Fault"(Core := #Core,
                   Status := #Status,
                   ReasonCode := 2021,
                   Description := WSTRING#'std.error.partCarrierWriteFailed');
       RETURN;
   END_IF;
   IF NOT "FRK_Carriers".Slots[#Index].Enabled THEN
       "FRK_Fault"(Core := #Core,
                   Status := #Status,
                   ReasonCode := 2021,
                   Description := WSTRING#'std.error.partCarrierWriteFailed');
       RETURN;
   END_IF;
   IF #Part.Uid <> "FRK_Carriers".Slots[#Index].Context.Uid THEN
       "FRK_Fault"(Core := #Core,
                   Status := #Status,
                   ReasonCode := 2022,
                   Description := WSTRING#'std.error.partCarrierReadFailed');
       RETURN;
   END_IF;
   #Part.Result.Verdict := #Verdict;
   #Part.Result.ReasonCode := #Reason;
   #Part.Result.StationPath := STRING_TO_WSTRING(#Status.Name);
   #Part.Result.TimeSynchronized := FALSE;
   #ResultCode := RD_SYS_T(OUT => #Stamp);
   IF #ResultCode = 0 THEN
       #Part.Result.Stamp := DTL_TO_LDT(#Stamp);
   END_IF;
   "FRK_Carriers".Slots[#Index].Written := #Part;
   IF "FRK_Carriers".Slots[#Index].Writes < UDINT#4294967295 THEN
       "FRK_Carriers".Slots[#Index].Writes := "FRK_Carriers".Slots[#Index].Writes + 1;
   END_IF;
   CASE #Verdict OF
       1:
           IF #Unit.Good < UDINT#4294967295 THEN
               #Unit.Good := #Unit.Good + 1;
           END_IF;
       2:
           IF #Unit.Nok < UDINT#4294967295 THEN
               #Unit.Nok := #Unit.Nok + 1;
           END_IF;
           #Unit.NokReason := #Reason;
       3:
           IF #Unit.Rework < UDINT#4294967295 THEN
               #Unit.Rework := #Unit.Rework + 1;
           END_IF;
       ELSE
           RETURN;
   END_CASE;
   // The provider result is written before publishing EVENT_PART_PROCESSED.
   "FRK_PartEvent"(AlarmLog := #AlarmLog,
                   Reason := 2026,
                   Uid := #Part.Uid,
                   SourcePath := #Status.Name);
   #Part.Present := FALSE;
   #FRK_PartProcessed := TRUE;
END_FUNCTION

FUNCTION "FRK_PartReceived" : Bool   // FC72, SCL
{ S7_Optimized_Access := 'TRUE' }
VERSION : 0.1
// stored: AutoNumber true, IsIECCheckEnabled false, SetENOAutomatically false, UDAEnableTagReadback false
   VAR_IN_OUT
      Core : "FRK_Core";
      Unit : "FRK_Unit";
      Status : "ST_ModuleStatus";
      Part : "ST_PartContext";
      AlarmLog : "FRK_AlarmLog";
   END_VAR
   VAR_TEMP
      Index : DInt;
      Uid : String[64];
      ResultIndex : DInt;
   END_VAR
BEGIN

   #FRK_PartReceived := FALSE;
   #Index := #Unit.CarrierIndex;
   IF #Index = 0 THEN
       RETURN;
   END_IF;
   IF #Index < 1 OR #Index > 32 THEN
       "FRK_Fault"(Core := #Core,
                   Status := #Status,
                   ReasonCode := 2020,
                   Description := WSTRING#'std.error.partCarrierReadFailed');
       RETURN;
   END_IF;
   IF NOT "FRK_Carriers".Slots[#Index].Enabled OR "FRK_Carriers".Slots[#Index].Kind <> 2 OR "FRK_Carriers".Slots[#Index].Serial = UDINT#4294967295 THEN
       "FRK_Fault"(Core := #Core,
                   Status := #Status,
                   ReasonCode := 2020,
                   Description := WSTRING#'std.error.partCarrierReadFailed');
       RETURN;
   END_IF;
   "FRK_Carriers".Slots[#Index].Serial := "FRK_Carriers".Slots[#Index].Serial + 1;
   #Uid := CONCAT(IN1 := 'FRK-', IN2 := DINT_TO_STRING(#Index));
   #Uid := CONCAT(IN1 := #Uid, IN2 := '-');
   #Uid := CONCAT(IN1 := #Uid, IN2 := UDINT_TO_STRING("FRK_Carriers".Slots[#Index].Serial));
   #Part.Uid := #Uid;
   #Part.Present := TRUE;
   #Part.CarrierKind := 2;
   #Part.Result.Verdict := 0;
   #Part.Result.ReasonCode := 0;
   #Part.Result.StationPath := STRING_TO_WSTRING(#Status.Name);
   #Part.Result.Stamp := LDT#1970-01-01-00:00:00.000000000;
   #Part.Result.TimeSynchronized := FALSE;
   FOR #ResultIndex := 1 TO 32 DO
       #Part.Result.Records[#ResultIndex].Name := '';
   END_FOR;
   FOR #ResultIndex := 1 TO 8 DO
       #Part.Parents[#ResultIndex] := '';
   END_FOR;
   "FRK_Carriers".Slots[#Index].Context := #Part;
   "FRK_PartEvent"(AlarmLog := #AlarmLog,
                   Reason := 2024,
                   Uid := #Part.Uid,
                   SourcePath := #Status.Name);
   #FRK_PartReceived := TRUE;
END_FUNCTION

FUNCTION "FRK_PartStarted" : Void   // FC73, SCL
{ S7_Optimized_Access := 'TRUE' }
VERSION : 0.1
// stored: AutoNumber true, IsIECCheckEnabled false, SetENOAutomatically false, UDAEnableTagReadback false
   VAR_IN_OUT
      Unit : "FRK_Unit";
      Status : "ST_ModuleStatus";
      Part : "ST_PartContext";
      AlarmLog : "FRK_AlarmLog";
   END_VAR
BEGIN

   IF #Unit.CarrierIndex = 0 OR NOT #Part.Present THEN
       RETURN;
   END_IF;
   "FRK_PartEvent"(AlarmLog := #AlarmLog,
                   Reason := 2025,
                   Uid := #Part.Uid,
                   SourcePath := #Status.Name);
END_FUNCTION

FUNCTION "FRK_PathOwned" : Bool   // FC86, SCL
{ S7_Optimized_Access := 'TRUE' }
VERSION : 0.1
// Shared Unit routing: typed generated edges carry these owning predicates.
// stored: AutoNumber true, IsIECCheckEnabled false, SetENOAutomatically false, UDAEnableTagReadback false
   VAR_INPUT
      OwnerPath : String;
      TargetPath : WString;
   END_VAR
   VAR_TEMP
      Width : Int;
   END_VAR
BEGIN

   #FRK_PathOwned := FALSE;
   #Width := LEN(#OwnerPath);
   IF #Width = 0 THEN
       RETURN;
   END_IF;
   IF #TargetPath = STRING_TO_WSTRING(#OwnerPath) THEN
       #FRK_PathOwned := TRUE;
       RETURN;
   END_IF;
   IF LEN(#TargetPath) <= #Width THEN
       RETURN;
   END_IF;
   #FRK_PathOwned := LEFT(IN := #TargetPath, L := #Width) = STRING_TO_WSTRING(#OwnerPath) AND #TargetPath[#Width + 1] = WCHAR#'.';
END_FUNCTION

FUNCTION "FRK_Pending" : Void   // FC13, SCL
{ S7_Optimized_Access := 'TRUE' }
VERSION : 0.1
// stored: AutoNumber true, IsIECCheckEnabled false, SetENOAutomatically false, UDAEnableTagReadback false
   VAR_INPUT
      Diag : "ST_Diagnostic";
   END_VAR
   VAR_IN_OUT
      Core : "FRK_Core";
      Status : "ST_ModuleStatus";
   END_VAR
BEGIN

   IF #Core.Exec = 1 AND NOT #Core.DiagTouched THEN
       #Status.Diagnostic := #Diag;
       #Status.Diagnostic.Severity := 0;
       #Core.DiagTouched := TRUE;
   END_IF;
END_FUNCTION

FUNCTION "FRK_Rationalize" : Void   // FC7, SCL
{ S7_Optimized_Access := 'TRUE' }
VERSION : 0.1
// stored: AutoNumber true, IsIECCheckEnabled false, SetENOAutomatically false, UDAEnableTagReadback false
   VAR_IN_OUT
      Diag : "ST_Diagnostic";
   END_VAR
BEGIN

   CASE #Diag.ReasonCode OF
       10:
           #Diag.Severity := 1;
           #Diag.Category := 2;
       11:
           #Diag.Severity := 0;
           #Diag.Category := 2;
       12:
           #Diag.Severity := 0;
           #Diag.Category := 2;
       13:
           #Diag.Severity := 1;
           #Diag.Category := 2;
       14:
           #Diag.Severity := 1;
           #Diag.Category := 2;
       15:
           #Diag.Severity := 2;
           #Diag.Category := 2;
       16:
           #Diag.Severity := 0;
           #Diag.Category := 2;
       17:
           #Diag.Severity := 0;
           #Diag.Category := 2;
       18:
           #Diag.Severity := 1;
           #Diag.Category := 2;
       19:
           #Diag.Severity := 0;
           #Diag.Category := 2;
       20:
           #Diag.Severity := 1;
           #Diag.Category := 2;
       21:
           #Diag.Severity := 0;
           #Diag.Category := 2;
       2001:
           #Diag.Severity := 1;
           #Diag.Category := 0;
       2002:
           #Diag.Severity := 0;
           #Diag.Category := 0;
       2003:
           #Diag.Severity := 1;
           #Diag.Category := 0;
       2004:
           #Diag.Severity := 1;
           #Diag.Category := 0;
       2005:
           #Diag.Severity := 0;
           #Diag.Category := 0;
       2006:
           #Diag.Severity := 1;
           #Diag.Category := 0;
       2007:
           #Diag.Severity := 0;
           #Diag.Category := 0;
       2008:
           #Diag.Severity := 0;
           #Diag.Category := 0;
       2010:
           #Diag.Severity := 1;
           #Diag.Category := 2;
       2011:
           #Diag.Severity := 0;
           #Diag.Category := 0;
       2012:
           #Diag.Severity := 1;
           #Diag.Category := 2;
       2020:
           #Diag.Severity := 1;
           #Diag.Category := 2;
       2021:
           #Diag.Severity := 1;
           #Diag.Category := 2;
       2022:
           #Diag.Severity := 2;
           #Diag.Category := 0;
       2023:
           #Diag.Severity := 1;
           #Diag.Category := 0;
       2024:
           #Diag.Severity := 0;
           #Diag.Category := 0;
       2025:
           #Diag.Severity := 0;
           #Diag.Category := 0;
       2026:
           #Diag.Severity := 0;
           #Diag.Category := 0;
       2027:
           #Diag.Severity := 0;
           #Diag.Category := 0;
       2030:
           #Diag.Severity := 0;
           #Diag.Category := 2;
       2040:
           #Diag.Severity := 1;
           #Diag.Category := 2;
       2041:
           #Diag.Severity := 1;
           #Diag.Category := 2;
       2042:
           #Diag.Severity := 0;
           #Diag.Category := 2;
       2043:
           #Diag.Severity := 0;
           #Diag.Category := 2;
       2901:
           #Diag.Severity := 0;
           #Diag.Category := 2;
       ELSE
           RETURN;
   END_CASE;
END_FUNCTION

FUNCTION "FRK_RecordTiming" : Void   // FC18, SCL
{ S7_Optimized_Access := 'TRUE' }
VERSION : 0.1
// stored: AutoNumber true, IsIECCheckEnabled false, SetENOAutomatically false, UDAEnableTagReadback false
   VAR_IN_OUT
      Core : "FRK_Core";
   END_VAR
   VAR_TEMP
      Index : DInt;
      Slot : DInt;
      DurationMs : UDInt;
      AverageMs : LInt;
   END_VAR
BEGIN

   #DurationMs := "FRK_Elapsed"(NewMs := "FRK_Clock".NowMs, OldMs := #Core.StartMs);
   // TIME's positive domain is bounded; clamp instead of publishing negatives.
   IF #DurationMs > UDINT#2147483647 THEN
       #DurationMs := UDINT#2147483647;
   END_IF;
   #Core.Timing.LastCmdTime := DINT_TO_TIME(UDINT_TO_DINT(#DurationMs));
   #Slot := 0;
   FOR #Index := 1 TO 8 DO
       IF #Core.Timing.Rows[#Index].Count > 0 AND #Core.Timing.Rows[#Index].Id = #Core.Command THEN
           #Slot := #Index;
           EXIT;
       ELSIF #Slot = 0 AND #Core.Timing.Rows[#Index].Count = 0 THEN
           #Slot := #Index;
       END_IF;
   END_FOR;
   IF #Slot = 0 THEN
       #Core.Timing.Truncated := TRUE;
   ELSE
       #Core.Timing.Rows[#Slot].Id := #Core.Command;
       #Core.Timing.Rows[#Slot].Label := #Core.CommandLabel;
       IF #Core.Timing.Rows[#Slot].Count < UDINT#4294967295 THEN
           #Core.Timing.Rows[#Slot].Count := #Core.Timing.Rows[#Slot].Count + 1;
       END_IF;
       #Core.Timing.Rows[#Slot].Last := #Core.Timing.LastCmdTime;
       IF #Core.Timing.Rows[#Slot].Count = 1 OR #Core.Timing.LastCmdTime < #Core.Timing.Rows[#Slot].Minimum THEN
           #Core.Timing.Rows[#Slot].Minimum := #Core.Timing.LastCmdTime;
       END_IF;
       IF #Core.Timing.LastCmdTime > #Core.Timing.Rows[#Slot].Maximum THEN
           #Core.Timing.Rows[#Slot].Maximum := #Core.Timing.LastCmdTime;
       END_IF;
       #AverageMs := DINT_TO_LINT(TIME_TO_DINT(#Core.Timing.Rows[#Slot].Avg));
       #AverageMs := #AverageMs + (UDINT_TO_LINT(#DurationMs) - #AverageMs) / UDINT_TO_LINT(#Core.Timing.Rows[#Slot].Count);
       #Core.Timing.Rows[#Slot].Avg := DINT_TO_TIME(LINT_TO_DINT(#AverageMs));
   END_IF;
   #Core.TimingOpen := FALSE;
END_FUNCTION

FUNCTION "FRK_ReleaseCommand" : Void   // FC20, SCL
{ S7_Optimized_Access := 'TRUE' }
VERSION : 0.1
// stored: AutoNumber true, IsIECCheckEnabled false, SetENOAutomatically false, UDAEnableTagReadback false
   VAR_IN_OUT
      Core : "FRK_Core";
      Execute : Bool;
   END_VAR
BEGIN

   #Execute := FALSE;
   #Core.ReleasePending := TRUE;
END_FUNCTION

FUNCTION "FRK_ReleaseReason" : Void   // FC77, SCL
{ S7_Optimized_Access := 'TRUE' }
VERSION : 0.1
// stored: AutoNumber true, IsIECCheckEnabled false, SetENOAutomatically false, UDAEnableTagReadback false
   VAR_INPUT
      Description : WString;
      Reason : DInt;
      Path : WString;
      Kind : DInt;
   END_VAR
   VAR_IN_OUT
      Report : "ST_ReleaseReport";
   END_VAR
BEGIN

   #Report.Released := FALSE;
   IF #Report.Count < 24 THEN
       #Report.Count := #Report.Count + 1;
       #Report.Reasons[#Report.Count].Description := #Description;
       #Report.Reasons[#Report.Count].ReasonCode := #Reason;
       #Report.Reasons[#Report.Count].SourcePath := #Path;
       #Report.Reasons[#Report.Count].Kind := #Kind;
       #Report.Reasons[#Report.Count].Bypassable := FALSE;
   END_IF;
END_FUNCTION

FUNCTION "FRK_Release_DeclarationUnit" : Void   // FC162, SCL
{ S7_Optimized_Access := 'TRUE' }
VERSION : 0.1
// stored: AutoNumber true, IsIECCheckEnabled false, SetENOAutomatically false, UDAEnableTagReadback false
   VAR_IN_OUT
      Unit : "FRK_Unit";
      Hal : "ST_DeclarationUnitHal";
   END_VAR
BEGIN

   "FRK_UnitSetPermit"(Unit := #Unit,
                       Ok := #Hal.Cell.Clamp.Permit,
                       Diag := #Hal.Cell.Clamp.Diag);
END_FUNCTION

FUNCTION "FRK_Release_InnerUnit" : Void   // FC146, SCL
{ S7_Optimized_Access := 'TRUE' }
VERSION : 0.1
// stored: AutoNumber true, IsIECCheckEnabled false, SetENOAutomatically false, UDAEnableTagReadback false
   VAR_IN_OUT
      Unit : "FRK_Unit";
      Hal : "ST_InnerUnitHal";
   END_VAR
BEGIN

   "FRK_UnitSetPermit"(Unit := #Unit,
                       Ok := #Hal.Cell.Clamp.Permit,
                       Diag := #Hal.Cell.Clamp.Diag);
END_FUNCTION

FUNCTION "FRK_Release_SatelliteUnit" : Void   // FC154, SCL
{ S7_Optimized_Access := 'TRUE' }
VERSION : 0.1
// stored: AutoNumber true, IsIECCheckEnabled false, SetENOAutomatically false, UDAEnableTagReadback false
   VAR_IN_OUT
      Unit : "FRK_Unit";
      Hal : "ST_SatelliteUnitHal";
   END_VAR
BEGIN

   "FRK_UnitSetPermit"(Unit := #Unit,
                       Ok := #Hal.Cell.Clamp.Permit,
                       Diag := #Hal.Cell.Clamp.Diag);
END_FUNCTION

FUNCTION "FRK_RouteAbort" : Void   // FC17, SCL
{ S7_Optimized_Access := 'TRUE' }
VERSION : 0.1
// stored: AutoNumber true, IsIECCheckEnabled false, SetENOAutomatically false, UDAEnableTagReadback false
   VAR_INPUT
      Abort : Bool;
   END_VAR
   VAR_IN_OUT
      Core : "FRK_Core";
   END_VAR
   VAR_TEMP
      ErrorAbort : Bool;
   END_VAR
BEGIN

   IF (#Abort OR #Core.ReleasePending) AND #Core.Exec = 1 THEN
       #Core.Exec := 4;
       #Core.Step := 0;
       #Core.Dispatch := FALSE;
       #Core.EvAbort := TRUE;
   END_IF;
   #ErrorAbort := (#Abort OR #Core.ReleasePending) AND #Core.Exec = 3;
   #Core.EvAbortInError := #ErrorAbort AND NOT #Core.AbortPrev;
   #Core.AbortPrev := #ErrorAbort;
END_FUNCTION

FUNCTION "FRK_Route_DeclarationCell" : Bool   // FC138, SCL
{ S7_Optimized_Access := 'TRUE' }
VERSION : 0.1
// stored: AutoNumber true, IsIECCheckEnabled false, SetENOAutomatically false, UDAEnableTagReadback false
   VAR_INPUT
      Request : "ST_HmiRequest";
   END_VAR
   VAR_IN_OUT
      Module : "FB_DeclarationCell";
      Hal : "ST_DeclarationCellHal";
      Report : "ST_ReleaseReport";
   END_VAR
   VAR_TEMP
      RouteMatched : Bool;
      Index : Int;
   END_VAR
BEGIN

